(* IEC 61131-3 sources: Industry-PLC-LLM/data/PLCBEAD_repo/PLCBEAD_PLCEmbed-main/PLC-BEAD/Source/PLC_Programs (part 7) *)

(* ---- GEN_RDT.ST ---- *)
FUNCTION _REAL_TO_UDINT:UDINT
  VAR_INPUT
    X :	REAL;
  END_VAR

  IF REAL_TO_UDINT(0.5) = UDINT#1 THEN
    _REAL_TO_UDINT := REAL_TO_UDINT(x);
  ELSIF X > 0.0 THEN
    _REAL_TO_UDINT := REAL_TO_UDINT(x+0.5);
  ELSIF X < 0.0 THEN
    _REAL_TO_UDINT := REAL_TO_UDINT(x-0.5);
  ELSE
    _REAL_TO_UDINT := UDINT#0;
  END_IF;
END_FUNCTION

FUNCTION REAL_TO_TIME2:TIME
	VAR_INPUT
		IN :	REAL;
	END_VAR

	REAL_TO_TIME2 := DINT_TO_TIME(UDINT_TO_DINT(_REAL_TO_UDINT(IN)));
END_FUNCTION

FUNCTION TIME_TO_REAL1:REAL

VAR_INPUT
	X :	TIME;
END_VAR

TIME_TO_REAL1 := UDINT_TO_REAL(DINT_TO_UDINT(TIME_TO_DINT(X)));
END_FUNCTION

FUNCTION D_TRUNC : DINT
  VAR_INPUT
    x : REAL;
  END_VAR

  D_TRUNC := REAL_TO_DINT(X);
  IF X > 0.0 THEN
  	IF DINT_TO_REAL(D_TRUNC) > X THEN D_TRUNC := D_TRUNC - DINT#1; END_IF;
  ELSE
  	IF DINT_TO_REAL(D_TRUNC) < X THEN D_TRUNC := D_TRUNC + DINT#1; END_IF;
  END_IF;
END_FUNCTION

FUNCTION BIT_COUNT:INT

	VAR_INPUT
		IN :	DWORD;
	END_VAR

	VAR
		in_temp :	DWORD;
	END_VAR

	in_temp := IN;
	WHILE in_temp > DWORD#0 DO
		IF (in_temp AND DWORD#16#00000001) > DWORD#0 THEN Bit_Count := Bit_Count +1; END_IF;
		in_temp := SHR(in_temp,1);
	END_WHILE;

END_FUNCTION

FUNCTION FRACT:REAL
	VAR_INPUT
		X :	REAL;
	END_VAR

	IF ABS(x) < 2.0E9 THEN
		FRACT := x - DINT_TO_REAL(D_TRUNC(x));
	ELSE
		FRACT := 0.0;
	END_IF;

END_FUNCTION

FUNCTION_BLOCK T_PLC_MS_block
	VAR_OUTPUT
		T_PLC_MS :	UDINT;
	END_VAR

	VAR_EXTERNAL
		PLC_TICKS_PER_SEC :	INT;
		PLC_SYS_TICK_CNT :	DINT;
	END_VAR

	VAR
		debug :	BOOL;(*Debug-Mode ON / OFF*)
		N :	INT;(*Debug-Faktor*)
		Offset :	UDINT;(*Debug-Offset*)
		temp :	DWORD := DWORD#1;(*Debug-Offset*)
		mode :	BOOL;(*modus*)
		faktor :	UDINT;(*Systemtakt-Faktor*)
		init :	BOOL;
		v_plc_ticks_per_sec :	UDINT;
		base :	UDINT := UDINT#1000;
	END_VAR

	IF init = FALSE THEN
		v_plc_ticks_per_sec := INT_TO_UDINT(PLC_TICKS_PER_SEC);
		IF v_plc_ticks_per_sec = UDINT#1024 THEN
			faktor := UDINT#1;
			mode := FALSE;
		ELSIF v_plc_ticks_per_sec > UDINT#0 THEN
			IF v_plc_ticks_per_sec <= base THEN
				faktor := base / v_plc_ticks_per_sec;
				mode := FALSE;
			ELSE
				faktor := v_plc_ticks_per_sec / base;
				mode := TRUE;
			END_IF;
		ELSE
			faktor := UDINT#1;
		END_IF;
		init := TRUE;
	END_IF;

	IF mode THEN
		T_PLC_MS := DINT_TO_UDINT(PLC_SYS_TICK_CNT) / faktor;
	ELSE
		T_PLC_MS := DINT_TO_UDINT(PLC_SYS_TICK_CNT) * faktor;
	END_IF;

	IF debug THEN
		T_PLC_MS := (DWORD_TO_UDINT(SHL(UDINT_TO_DWORD(T_PLC_MS),N) OR SHL(temp,N)) - UDINT#1) + Offset;
	END_IF;

END_FUNCTION_BLOCK

FUNCTION BIT_LOAD_DW:DWORD

	VAR_INPUT
		IN :	DWORD;
		VAL :	BOOL;
		POS :	INT;
	END_VAR

	IF val THEN
		BIT_LOAD_DW := in OR SHL(DWORD#1,pos);
	ELSE
		BIT_LOAD_DW := in AND (NOT SHL(DWORD#1,pos));
	END_IF;

END_FUNCTION

FUNCTION BIT_OF_DWORD : BOOL
  VAR_INPUT
    IN : DWORD;
    N : INT;
  END_VAR

  BIT_OF_DWORD := (SHR(in,N) AND 16#00000001) > 0;
  (* from OSCAT library; www.oscat.de  *)
END_FUNCTION

FUNCTION _INT_TO_UDINT:UDINT
	VAR_INPUT
		IN :	INT;
	END_VAR

	_INT_TO_UDINT := DINT_TO_UDINT(INT_TO_DINT(IN));
END_FUNCTION

FUNCTION _DWORD_TO_REAL:REAL
	VAR_INPUT
		IN :	DWORD;
	END_VAR

	_DWORD_TO_REAL := UDINT_TO_REAL(DWORD_TO_UDINT(IN));

END_FUNCTION

FUNCTION_BLOCK RDM_block
	VAR_INPUT
		LAST :	REAL;
	END_VAR
	VAR_OUTPUT
		RDM :	REAL;
	END_VAR
	VAR
		T_PLC_MS :	T_PLC_MS_block;
		tn :	DWORD;
		tc :	INT;
	END_VAR
	T_PLC_MS();
	tn := UDINT_TO_DWORD(T_PLC_MS.T_PLC_MS);
	tc := Bit_Count(tn);

	tn:=BIT_LOAD_DW(tn,BIT_OF_DWORD(tn,2),31); (* tn.31 := tn.2; *)
	tn:=BIT_LOAD_DW(tn,BIT_OF_DWORD(tn,5),30); (* tn.30 := tn.5; *)
	tn:=BIT_LOAD_DW(tn,BIT_OF_DWORD(tn,4),29); (* tn.29 := tn.4; *)
	tn:=BIT_LOAD_DW(tn,BIT_OF_DWORD(tn,1),28); (* tn.28 := tn.1; *)
	tn:=BIT_LOAD_DW(tn,BIT_OF_DWORD(tn,0),27); (* tn.27 := tn.0; *)
	tn:=BIT_LOAD_DW(tn,BIT_OF_DWORD(tn,7),26); (* tn.26 := tn.7; *)
	tn:=BIT_LOAD_DW(tn,BIT_OF_DWORD(tn,6),25); (* tn.25 := tn.6; *)
	tn:=BIT_LOAD_DW(tn,BIT_OF_DWORD(tn,3),24); (* tn.24 := tn.3; *)

	tn := ROL(tn,Bit_Count(tn)) OR DWORD#16#80000001;
	tn := UDINT_TO_DWORD(DWORD_TO_UDINT(tn) MOD UDINT#71474513 + _INT_TO_UDINT(tc) + UDINT#77);
	RDM := fract(_DWORD_TO_REAL(tn) / 10000000.0 * (2.71828182845904523536028747135266249 - LIMIT_REAL(0.0,last,1.0)));
END_FUNCTION_BLOCK

FUNCTION_BLOCK GEN_RDT_Block

	VAR_INPUT
		ENABLE :	BOOL := TRUE;
		MIN_TIME_MS :	TIME := t#1s;
		MAX_TIME_MS :	TIME := t#1.2s;
		TP_Q :	TIME := t#100ms;
	END_VAR

	VAR_OUTPUT
		XQ :	BOOL;
	END_VAR

	VAR
		tonRDMTimer :	TON;
		tof_xQ :	TOF;
		tRDMTime :	TIME;
		rRDMTime :	REAL;
		rdm_1 :	RDM_Block;
	END_VAR

	tonRDMTimer(IN:=Enable,PT:=tRDMTime);
	tof_xQ(IN := tonRDMTimer.Q,PT:=TP_Q);
	XQ := tof_xq.Q;
	IF tonRDMTimer.Q THEN
		xQ := TRUE ;
		rdm_1(last:=rRDMTime);
		rRDMTime:= rdm_1.RDM;

		tRDMTime := REAL_TO_TIME2(rRDMTime * TIME_TO_REAL1(Max_Time_ms - Min_Time_ms) + TIME_TO_REAL1(Min_Time_ms));
		tonRDMTimer (IN:=FALSE);
	END_IF;

END_FUNCTION_BLOCK

PROGRAM program0
  VAR
	ENABLE :	BOOL := TRUE;
	MIN_TIME_MS :	TIME := t#1s;
	MAX_TIME_MS :	TIME := t#1.2s;
	TP_Q :	TIME := t#100ms;
	XQ :	BOOL;
	func_block : GEN_RDT_Block;
  END_VAR
	func_block.ENABLE  :=ENABLE;
	func_block.MIN_TIME_MS  :=MIN_TIME_MS;
	func_block.MAX_TIME_MS  :=MAX_TIME_MS;
	func_block.TP_Q  :=TP_Q;
	func_block();
	XQ := func_block.XQ;
END_PROGRAM

CONFIGURATION Config0
	VAR_GLOBAL
		PLC_TICKS_PER_SEC :	INT;
		PLC_SYS_TICK_CNT :	DINT;
	END_VAR
	RESOURCE Res0 ON PLC
		TASK task0(INTERVAL := T#20ms,PRIORITY := 0);
		PROGRAM instance0 WITH task0 : program0;
	END_RESOURCE
END_CONFIGURATION

(* ---- GEN_RMP.ST ---- *)
FUNCTION D_TRUNC : DINT
  VAR_INPUT
    x : REAL;
  END_VAR

  D_TRUNC := REAL_TO_DINT(X);
  IF X > 0.0 THEN
  	IF DINT_TO_REAL(D_TRUNC) > X THEN D_TRUNC := D_TRUNC - DINT#1; END_IF;
  ELSE
  	IF DINT_TO_REAL(D_TRUNC) < X THEN D_TRUNC := D_TRUNC + DINT#1; END_IF;
  END_IF;
END_FUNCTION

FUNCTION FRACT:REAL
	VAR_INPUT
		X :	REAL;
	END_VAR

	IF ABS(x) < 2.0E9 THEN
		FRACT := x - DINT_TO_REAL(D_TRUNC(x));
	ELSE
		FRACT := 0.0;
	END_IF;
END_FUNCTION

FUNCTION _REAL_TO_DWORD: DWORD

  VAR_INPUT
    X :	REAL;
  END_VAR

  IF REAL_TO_DWORD(0.5) = DWORD#1 THEN
    _REAL_TO_DWORD := REAL_TO_DWORD(x);
  ELSIF X > 0.0 THEN
    _REAL_TO_DWORD := REAL_TO_DWORD(x+0.5);
  ELSIF X < 0.0 THEN
    _REAL_TO_DWORD := REAL_TO_DWORD(x-0.5);
  ELSE
    _REAL_TO_DWORD := DWORD#0;
  END_IF;
END_FUNCTION

FUNCTION _DWORD_TO_REAL:REAL
	VAR_INPUT
		IN :	DWORD;
	END_VAR

	_DWORD_TO_REAL := UDINT_TO_REAL(DWORD_TO_UDINT(IN));

END_FUNCTION

FUNCTION MULTIME:TIME
	VAR_INPUT
		T :	TIME;
		M :	REAL;
	END_VAR

	multime := DWORD_TO_TIME(_REAL_TO_DWORD(_DWORD_TO_REAL(TIME_TO_DWORD(t))*M));
END_FUNCTION

FUNCTION TIME_TO_REAL1:REAL

VAR_INPUT
	X :	TIME;
END_VAR

TIME_TO_REAL1 := UDINT_TO_REAL(DINT_TO_UDINT(TIME_TO_DINT(X)));
END_FUNCTION

FUNCTION MODR : REAL
  VAR_INPUT
    IN : REAL;
    DIVI : REAL;
  END_VAR

  IF divi = 0.0 THEN
  	MODR := 0.0;
  ELSE
  	MODR := in - DINT_TO_REAL(FLOOR2(in / divi)) * divi;
  END_IF;
END_FUNCTION

FUNCTION FLOOR2 : DINT
  VAR_INPUT
    x : REAL;
  END_VAR

  FLOOR2 := REAL_TO_DINT(X);
  IF DINT_TO_REAL(FLOOR2) > X THEN
  	FLOOR2 := FLOOR2 - DINT#1;
  END_IF;
END_FUNCTION

FUNCTION UDINT_TO_TIME2:TIME

	VAR_INPUT
		IN :	UDINT;
	END_VAR

	UDINT_TO_TIME2 := DINT_TO_TIME(UDINT_TO_DINT(IN));

END_FUNCTION

FUNCTION_BLOCK T_PLC_MS_block
	VAR_OUTPUT
		T_PLC_MS :	UDINT;
	END_VAR

	VAR_EXTERNAL
		PLC_TICKS_PER_SEC :	INT;
		PLC_SYS_TICK_CNT :	DINT;
	END_VAR

	VAR
		debug :	BOOL;(*Debug-Mode ON / OFF*)
		N :	INT;(*Debug-Faktor*)
		Offset :	UDINT;(*Debug-Offset*)
		temp :	DWORD := DWORD#1;(*Debug-Offset*)
		mode :	BOOL;(*modus*)
		faktor :	UDINT;(*Systemtakt-Faktor*)
		init :	BOOL;
		v_plc_ticks_per_sec :	UDINT;
		base :	UDINT := UDINT#1000;
	END_VAR

	IF init = FALSE THEN
		v_plc_ticks_per_sec := INT_TO_UDINT(PLC_TICKS_PER_SEC);
		IF v_plc_ticks_per_sec = UDINT#1024 THEN
			faktor := UDINT#1;
			mode := FALSE;
		ELSIF v_plc_ticks_per_sec > UDINT#0 THEN
			IF v_plc_ticks_per_sec <= base THEN
				faktor := base / v_plc_ticks_per_sec;
				mode := FALSE;
			ELSE
				faktor := v_plc_ticks_per_sec / base;
				mode := TRUE;
			END_IF;
		ELSE
			faktor := UDINT#1;
		END_IF;
		init := TRUE;
	END_IF;

	IF mode THEN
		T_PLC_MS := DINT_TO_UDINT(PLC_SYS_TICK_CNT) / faktor;
	ELSE
		T_PLC_MS := DINT_TO_UDINT(PLC_SYS_TICK_CNT) * faktor;
	END_IF;

	IF debug THEN
		T_PLC_MS := (DWORD_TO_UDINT(SHL(UDINT_TO_DWORD(T_PLC_MS),N) OR SHL(temp,N)) - UDINT#1) + Offset;
	END_IF;

END_FUNCTION_BLOCK

FUNCTION_BLOCK GEN_RMP_Block

	VAR_INPUT
		PT :	TIME := T#1s;
		AM :	REAL := REAL#1.0;
		OS :	REAL;
		DL :	REAL;
	END_VAR

	VAR_OUTPUT
		Q :	BOOL;
		OUT :	REAL;
	END_VAR

	VAR
		tx :	TIME;
		last :	TIME;
		init :	BOOL;
		temp :	REAL;
		ltemp :	REAL;
		T_PLC_MS :	T_PLC_MS_Block;
	END_VAR

	T_PLC_MS();
	tx:= UDINT_TO_TIME(T_PLC_MS.T_PLC_MS) - last;
	DL := modR(dl,1.0);
	IF dl < 0.0 THEN dl := 1.0 - dl; END_IF;

	IF NOT init THEN
		init := TRUE;
		last := tx;
		tx := t#0s;
	END_IF;

	IF tx >= pt THEN
		last := last + pt;
		tx := tx - pt;
	END_IF;

	ltemp := temp;
	IF pt > t#0s THEN temp := fract(TIME_TO_REAL1(tx + multime(pt, dl)) / TIME_TO_REAL1(pt)); END_IF;
	out := am * temp + os;

	Q := temp < ltemp;

END_FUNCTION_BLOCK

PROGRAM program0
  VAR
	PT :	TIME := T#1s;
	AM :	REAL := REAL#1.0;
	OS :	REAL;
	DL :	REAL;
	Q :	BOOL;
	OUT :	REAL;
	func_block : GEN_RMP_Block;
  END_VAR
	func_block.PT  :=PT;
	func_block.AM  :=AM;
	func_block.OS  :=OS;
	func_block.DL  :=DL;
	func_block();
	Q := func_block.Q;
	OUT := func_block.OUT;
END_PROGRAM

CONFIGURATION Config0
	VAR_GLOBAL
		PLC_TICKS_PER_SEC :	INT;
		PLC_SYS_TICK_CNT :	DINT;
	END_VAR
	RESOURCE Res0 ON PLC
		TASK task0(INTERVAL := T#20ms,PRIORITY := 0);
		PROGRAM instance0 WITH task0 : program0;
	END_RESOURCE
END_CONFIGURATION

(* ---- GEN_SIN.ST ---- *)
FUNCTION _REAL_TO_DWORD: DWORD

  VAR_INPUT
    X :	REAL;
  END_VAR

  IF REAL_TO_DWORD(0.5) = DWORD#1 THEN
    _REAL_TO_DWORD := REAL_TO_DWORD(x);
  ELSIF X > 0.0 THEN
    _REAL_TO_DWORD := REAL_TO_DWORD(x+0.5);
  ELSIF X < 0.0 THEN
    _REAL_TO_DWORD := REAL_TO_DWORD(x-0.5);
  ELSE
    _REAL_TO_DWORD := DWORD#0;
  END_IF;
END_FUNCTION

FUNCTION _DWORD_TO_REAL:REAL
	VAR_INPUT
		IN :	DWORD;
	END_VAR

	_DWORD_TO_REAL := UDINT_TO_REAL(DWORD_TO_UDINT(IN));

END_FUNCTION

FUNCTION MULTIME:TIME
	VAR_INPUT
		T :	TIME;
		M :	REAL;
	END_VAR

	multime := DWORD_TO_TIME(_REAL_TO_DWORD(_DWORD_TO_REAL(TIME_TO_DWORD(t))*M));
END_FUNCTION

FUNCTION UDINT_TO_TIME2:TIME

	VAR_INPUT
		IN :	UDINT;
	END_VAR

	UDINT_TO_TIME2 := DINT_TO_TIME(UDINT_TO_DINT(IN));

END_FUNCTION

FUNCTION_BLOCK T_PLC_MS_block
	VAR_OUTPUT
		T_PLC_MS :	UDINT;
	END_VAR

	VAR_EXTERNAL
		PLC_TICKS_PER_SEC :	INT;
		PLC_SYS_TICK_CNT :	DINT;
	END_VAR

	VAR
		debug :	BOOL;(*Debug-Mode ON / OFF*)
		N :	INT;(*Debug-Faktor*)
		Offset :	UDINT;(*Debug-Offset*)
		temp :	DWORD := DWORD#1;(*Debug-Offset*)
		mode :	BOOL;(*modus*)
		faktor :	UDINT;(*Systemtakt-Faktor*)
		init :	BOOL;
		v_plc_ticks_per_sec :	UDINT;
		base :	UDINT := UDINT#1000;
	END_VAR

	IF init = FALSE THEN
		v_plc_ticks_per_sec := INT_TO_UDINT(PLC_TICKS_PER_SEC);
		IF v_plc_ticks_per_sec = UDINT#1024 THEN
			faktor := UDINT#1;
			mode := FALSE;
		ELSIF v_plc_ticks_per_sec > UDINT#0 THEN
			IF v_plc_ticks_per_sec <= base THEN
				faktor := base / v_plc_ticks_per_sec;
				mode := FALSE;
			ELSE
				faktor := v_plc_ticks_per_sec / base;
				mode := TRUE;
			END_IF;
		ELSE
			faktor := UDINT#1;
		END_IF;
		init := TRUE;
	END_IF;

	IF mode THEN
		T_PLC_MS := DINT_TO_UDINT(PLC_SYS_TICK_CNT) / faktor;
	ELSE
		T_PLC_MS := DINT_TO_UDINT(PLC_SYS_TICK_CNT) * faktor;
	END_IF;

	IF debug THEN
		T_PLC_MS := (DWORD_TO_UDINT(SHL(UDINT_TO_DWORD(T_PLC_MS),N) OR SHL(temp,N)) - UDINT#1) + Offset;
	END_IF;

END_FUNCTION_BLOCK

FUNCTION TIME_TO_REAL1:REAL

	VAR_INPUT
		X :	TIME;
	END_VAR

	TIME_TO_REAL1 := UDINT_TO_REAL(DINT_TO_UDINT(TIME_TO_DINT(X)));
END_FUNCTION

FUNCTION MODR : REAL
  VAR_INPUT
    IN : REAL;
    DIVI : REAL;
  END_VAR

  IF divi = 0.0 THEN
  	MODR := 0.0;
  ELSE
  	MODR := in - DINT_TO_REAL(FLOOR2(in / divi)) * divi;
  END_IF;
END_FUNCTION

FUNCTION FLOOR2 : DINT
  VAR_INPUT
    x : REAL;
  END_VAR

  FLOOR2 := REAL_TO_DINT(X);
  IF DINT_TO_REAL(FLOOR2) > X THEN
  	FLOOR2 := FLOOR2 - DINT#1;
  END_IF;
END_FUNCTION

FUNCTION SIGN_R : BOOL
  VAR_INPUT
    IN : REAL;
  END_VAR

  SIGN_R := in < 0.0;
END_FUNCTION

FUNCTION_BLOCK GEN_SIN_Block

	VAR_INPUT
		PT :	TIME;
		AM :	REAL := REAL#1.0;
		OS :	REAL;
		DL :	REAL;
	END_VAR

	VAR_OUTPUT
		Q :	BOOL;
		Out :	REAL;
	END_VAR

	VAR
		tx :	TIME;
		last :	TIME;
		init :	BOOL;
		temp :	REAL;
		T_PLC_MS :	T_PLC_MS_Block;
	END_VAR

	T_PLC_MS();
	tx:= UDINT_TO_TIME(T_PLC_MS.T_PLC_MS) - last;

	DL := modR(dl,1.0);
	IF dl < 0.0 THEN dl := 1.0 - dl; END_IF;

	IF NOT init THEN
		init := TRUE;
		last := tx;
		tx := t#0s;
	END_IF;

	IF tx >= pt THEN
		last := last + pt;
		tx := tx - pt;
	END_IF;

	IF pt > t#0s THEN temp := SIN(6.283185307179586476 * TIME_TO_REAL1(tx + multime(pt, dl)) / TIME_TO_REAL(pt)); END_IF;
	out := am * 0.5 *  temp + os;

	q := NOT sign_R(temp);

END_FUNCTION_BLOCK

PROGRAM program0
  VAR
	PT :	TIME := T#1s;
	AM :	REAL := REAL#1.0;
	OS :	REAL;
	DL :	REAL;
	Q :	BOOL;
	OUT :	REAL;
	func_block : GEN_SIN_Block;
  END_VAR
	func_block.PT  :=PT;
	func_block.AM  :=AM;
	func_block.OS  :=OS;
	func_block.DL  :=DL;
	func_block();
	Q := func_block.Q;
	OUT := func_block.OUT;
END_PROGRAM

CONFIGURATION Config0
	VAR_GLOBAL
		PLC_TICKS_PER_SEC :	INT;
		PLC_SYS_TICK_CNT :	DINT;
	END_VAR
	RESOURCE Res0 ON PLC
		TASK task0(INTERVAL := T#20ms,PRIORITY := 0);
		PROGRAM instance0 WITH task0 : program0;
	END_RESOURCE
END_CONFIGURATION

(* ---- GEN_SQ.ST ---- *)
FUNCTION UDINT_TO_TIME2:TIME

	VAR_INPUT
		IN :	UDINT;
	END_VAR

	UDINT_TO_TIME2 := DINT_TO_TIME(UDINT_TO_DINT(IN));

END_FUNCTION

FUNCTION_BLOCK T_PLC_MS_block
	VAR_OUTPUT
		T_PLC_MS :	UDINT;
	END_VAR

	VAR_EXTERNAL
		PLC_TICKS_PER_SEC :	INT;
		PLC_SYS_TICK_CNT :	DINT;
	END_VAR

	VAR
		debug :	BOOL;(*Debug-Mode ON / OFF*)
		N :	INT;(*Debug-Faktor*)
		Offset :	UDINT;(*Debug-Offset*)
		temp :	DWORD := DWORD#1;(*Debug-Offset*)
		mode :	BOOL;(*modus*)
		faktor :	UDINT;(*Systemtakt-Faktor*)
		init :	BOOL;
		v_plc_ticks_per_sec :	UDINT;
		base :	UDINT := UDINT#1000;
	END_VAR

	IF init = FALSE THEN
		v_plc_ticks_per_sec := INT_TO_UDINT(PLC_TICKS_PER_SEC);
		IF v_plc_ticks_per_sec = UDINT#1024 THEN
			faktor := UDINT#1;
			mode := FALSE;
		ELSIF v_plc_ticks_per_sec > UDINT#0 THEN
			IF v_plc_ticks_per_sec <= base THEN
				faktor := base / v_plc_ticks_per_sec;
				mode := FALSE;
			ELSE
				faktor := v_plc_ticks_per_sec / base;
				mode := TRUE;
			END_IF;
		ELSE
			faktor := UDINT#1;
		END_IF;
		init := TRUE;
	END_IF;

	IF mode THEN
		T_PLC_MS := DINT_TO_UDINT(PLC_SYS_TICK_CNT) / faktor;
	ELSE
		T_PLC_MS := DINT_TO_UDINT(PLC_SYS_TICK_CNT) * faktor;
	END_IF;

	IF debug THEN
		T_PLC_MS := (DWORD_TO_UDINT(SHL(UDINT_TO_DWORD(T_PLC_MS),N) OR SHL(temp,N)) - UDINT#1) + Offset;
	END_IF;

END_FUNCTION_BLOCK

FUNCTION_BLOCK GEN_SQ_Block

	VAR_INPUT
		PT :	TIME;
	END_VAR

	VAR_OUTPUT
		Q :	BOOL;
	END_VAR

	VAR
		init :	BOOL;
		tn :	TIME;
		tx :	TIME;
		T_PLC_MS :	T_PLC_MS_Block;
	END_VAR

	T_PLC_MS();
	tx := UDINT_TO_TIME(T_PLC_MS.T_PLC_MS);

	IF NOT init THEN
		init := TRUE;
		tn := tx;
		Q := TRUE;
	ELSIF tx - tn >= DWORD_TO_TIME(SHR(TIME_TO_DWORD(PT),1)) THEN
		Q := NOT Q;
		tn := tn + DWORD_TO_TIME(SHR(TIME_TO_DWORD(pt),1));
	END_IF;

END_FUNCTION_BLOCK

PROGRAM program0
  VAR
	PT :	TIME;
	Q :	BOOL;
	OUT :	REAL;
	func_block : GEN_SQ_Block;
  END_VAR
	func_block.PT  :=PT;
	func_block();
	Q := func_block.Q;
END_PROGRAM

CONFIGURATION Config0
	VAR_GLOBAL
		PLC_TICKS_PER_SEC :	INT;
		PLC_SYS_TICK_CNT :	DINT;
	END_VAR
	RESOURCE Res0 ON PLC
		TASK task0(INTERVAL := T#20ms,PRIORITY := 0);
		PROGRAM instance0 WITH task0 : program0;
	END_RESOURCE
END_CONFIGURATION

(* ---- GEN_SQR.ST ---- *)
FUNCTION UDINT_TO_TIME2:TIME

	VAR_INPUT
		IN :	UDINT;
	END_VAR

	UDINT_TO_TIME2 := DINT_TO_TIME(UDINT_TO_DINT(IN));

END_FUNCTION

FUNCTION_BLOCK T_PLC_MS_block
	VAR_OUTPUT
		T_PLC_MS :	UDINT;
	END_VAR

	VAR_EXTERNAL
		PLC_TICKS_PER_SEC :	INT;
		PLC_SYS_TICK_CNT :	DINT;
	END_VAR

	VAR
		debug :	BOOL;(*Debug-Mode ON / OFF*)
		N :	INT;(*Debug-Faktor*)
		Offset :	UDINT;(*Debug-Offset*)
		temp :	DWORD := DWORD#1;(*Debug-Offset*)
		mode :	BOOL;(*modus*)
		faktor :	UDINT;(*Systemtakt-Faktor*)
		init :	BOOL;
		v_plc_ticks_per_sec :	UDINT;
		base :	UDINT := UDINT#1000;
	END_VAR

	IF init = FALSE THEN
		v_plc_ticks_per_sec := INT_TO_UDINT(PLC_TICKS_PER_SEC);
		IF v_plc_ticks_per_sec = UDINT#1024 THEN
			faktor := UDINT#1;
			mode := FALSE;
		ELSIF v_plc_ticks_per_sec > UDINT#0 THEN
			IF v_plc_ticks_per_sec <= base THEN
				faktor := base / v_plc_ticks_per_sec;
				mode := FALSE;
			ELSE
				faktor := v_plc_ticks_per_sec / base;
				mode := TRUE;
			END_IF;
		ELSE
			faktor := UDINT#1;
		END_IF;
		init := TRUE;
	END_IF;

	IF mode THEN
		T_PLC_MS := DINT_TO_UDINT(PLC_SYS_TICK_CNT) / faktor;
	ELSE
		T_PLC_MS := DINT_TO_UDINT(PLC_SYS_TICK_CNT) * faktor;
	END_IF;

	IF debug THEN
		T_PLC_MS := (DWORD_TO_UDINT(SHL(UDINT_TO_DWORD(T_PLC_MS),N) OR SHL(temp,N)) - UDINT#1) + Offset;
	END_IF;

END_FUNCTION_BLOCK

FUNCTION MODR : REAL
  VAR_INPUT
    IN : REAL;
    DIVI : REAL;
  END_VAR

  IF divi = 0.0 THEN
  	MODR := 0.0;
  ELSE
  	MODR := in - DINT_TO_REAL(FLOOR2(in / divi)) * divi;
  END_IF;
END_FUNCTION

FUNCTION FLOOR2 : DINT
  VAR_INPUT
    x : REAL;
  END_VAR

  FLOOR2 := REAL_TO_DINT(X);
  IF DINT_TO_REAL(FLOOR2) > X THEN
  	FLOOR2 := FLOOR2 - DINT#1;
  END_IF;
END_FUNCTION

FUNCTION _REAL_TO_DWORD: DWORD

  VAR_INPUT
    X :	REAL;
  END_VAR

  IF REAL_TO_DWORD(0.5) = DWORD#1 THEN
    _REAL_TO_DWORD := REAL_TO_DWORD(x);
  ELSIF X > 0.0 THEN
    _REAL_TO_DWORD := REAL_TO_DWORD(x+0.5);
  ELSIF X < 0.0 THEN
    _REAL_TO_DWORD := REAL_TO_DWORD(x-0.5);
  ELSE
    _REAL_TO_DWORD := DWORD#0;
  END_IF;
END_FUNCTION

FUNCTION _DWORD_TO_REAL:REAL
	VAR_INPUT
		IN :	DWORD;
	END_VAR

	_DWORD_TO_REAL := UDINT_TO_REAL(DWORD_TO_UDINT(IN));

END_FUNCTION

FUNCTION MULTIME:TIME
	VAR_INPUT
		T :	TIME;
		M :	REAL;
	END_VAR

	multime := DWORD_TO_TIME(_REAL_TO_DWORD(_DWORD_TO_REAL(TIME_TO_DWORD(t))*M));
END_FUNCTION

FUNCTION_BLOCK GEN_SQR_Block

	VAR_INPUT
		PT :	TIME;
		AM :	REAL := REAL#1.0;
		OS :	REAL;
		DC :	REAL := REAL#0.5;
		DL :	REAL;
	END_VAR

	VAR_OUTPUT
		Q :	BOOL;
		Out :	REAL;
	END_VAR

	VAR
		tx :	TIME;
		last :	TIME;
		init :	BOOL;
		T_PLC_MS :	T_PLC_MS_Block;
	END_VAR

	IF dc = 0.0 THEN
		out := -am * 0.5 + os;
		Q := FALSE;
		RETURN;
	ELSIF dc = 1.0 THEN
		out := am * 0.5 + os;
		Q := TRUE;
		RETURN;
	END_IF;

	T_PLC_MS();
	tx:= UDINT_TO_TIME(T_PLC_MS.T_PLC_MS) - last;
	DL := modR(dl,1.0);
	IF dl < 0.0 THEN dl := 1.0 - dl; END_IF;
	dc := modR(dc,1.0);
	IF dc < 0.0 THEN dc := 1.0 - dc; END_IF;

	IF NOT init THEN
		init := TRUE;
		last := tx;
		tx := t#0s;
	END_IF;

	IF tx >= pt THEN
		last := last + pt;
		tx := tx - pt;
	END_IF;

	IF multime(pt, dl + dc) >= pt THEN
		IF tx >= multime(pt, dl + dc - 1.0) THEN
			out := -am * 0.5 + os;
			Q := FALSE;
		END_IF;
		IF tx >= multime(pt, dl) THEN
			out := am * 0.5 + os;
			Q := TRUE;
		END_IF;
	ELSE
		IF tx >= multime(pt, dl) THEN
			out := am * 0.5 + os;
			Q := TRUE;
		END_IF;
		IF tx >= multime(pt, dl + dc) THEN
			out := -am * 0.5 +os;
			Q := FALSE;
		END_IF;
	END_IF;

END_FUNCTION_BLOCK

PROGRAM program0
  VAR
	PT :	TIME;
	AM :	REAL := REAL#1.0;
	OS :	REAL;
	DC :	REAL := REAL#0.5;
	DL :	REAL;
	Q :	BOOL;
	Out :	REAL;
	func_block : GEN_SQR_Block;
  END_VAR
	func_block.PT  :=PT;
	func_block.AM  :=AM;
	func_block.OS  :=OS;
	func_block.DC  :=DC;
	func_block.DL  :=DL;
	func_block();
	Q := func_block.Q;
	OUT := func_block.OUT;
END_PROGRAM

CONFIGURATION Config0
	VAR_GLOBAL
		PLC_TICKS_PER_SEC :	INT;
		PLC_SYS_TICK_CNT :	DINT;
	END_VAR
	RESOURCE Res0 ON PLC
		TASK task0(INTERVAL := T#20ms,PRIORITY := 0);
		PROGRAM instance0 WITH task0 : program0;
	END_RESOURCE
END_CONFIGURATION

(* ---- HEAT_METER.ST ---- *)
FUNCTION UDINT_TO_TIME2:TIME
	VAR_INPUT
		IN :	UDINT;
	END_VAR
	UDINT_TO_TIME2 := DINT_TO_TIME(UDINT_TO_DINT(IN));
END_FUNCTION

FUNCTION_BLOCK T_PLC_MS_block
	VAR_OUTPUT
		T_PLC_MS :	UDINT;
	END_VAR

	VAR_EXTERNAL
		PLC_TICKS_PER_SEC :	INT;
		PLC_SYS_TICK_CNT :	DINT;
	END_VAR

	VAR
		debug :	BOOL;(*Debug-Mode ON / OFF*)
		N :	INT;(*Debug-Faktor*)
		Offset :	UDINT;(*Debug-Offset*)
		temp :	DWORD := DWORD#1;(*Debug-Offset*)
		mode :	BOOL;(*modus*)
		faktor :	UDINT;(*Systemtakt-Faktor*)
		init :	BOOL;
		v_plc_ticks_per_sec :	UDINT;
		base :	UDINT := UDINT#1000;
	END_VAR

	IF init = FALSE THEN
		v_plc_ticks_per_sec := INT_TO_UDINT(PLC_TICKS_PER_SEC);
		IF v_plc_ticks_per_sec = UDINT#1024 THEN
			faktor := UDINT#1;
			mode := FALSE;
		ELSIF v_plc_ticks_per_sec > UDINT#0 THEN
			IF v_plc_ticks_per_sec <= base THEN
				faktor := base / v_plc_ticks_per_sec;
				mode := FALSE;
			ELSE
				faktor := v_plc_ticks_per_sec / base;
				mode := TRUE;
			END_IF;
		ELSE
			faktor := UDINT#1;
		END_IF;
		init := TRUE;
	END_IF;

	IF mode THEN
		T_PLC_MS := DINT_TO_UDINT(PLC_SYS_TICK_CNT) / faktor;
	ELSE
		T_PLC_MS := DINT_TO_UDINT(PLC_SYS_TICK_CNT) * faktor;
	END_IF;

	IF debug THEN
		T_PLC_MS := (DWORD_TO_UDINT(SHL(UDINT_TO_DWORD(T_PLC_MS),N) OR SHL(temp,N)) - UDINT#1) + Offset;
	END_IF;

END_FUNCTION_BLOCK

TYPE
	oscat_ARRAY_X               : ARRAY [0..1]    OF REAL;
	oscat_XY                    : ARRAY [1..20]   OF oscat_ARRAY_X := [0,0,0,0,0,0,0,0,0,0,0,0,0,0,0,0,0,0,0,0];
END_TYPE

FUNCTION_BLOCK LINEAR_INT_Block

	VAR_INPUT
		X :	REAL;
		XY :	oscat_XY;
		PTS :	INT;
	END_VAR

	VAR_OUTPUT
		LINEAR_INT :	REAL;
	END_VAR

	VAR
		i :	INT;
		i2 :	INT;
	END_VAR

	pts := MIN(pts,20);

	i := 2;

	WHILE (i < pts) AND (XY[i][0] < X) DO
		i := i + 1;
	END_WHILE;

	i2 := i-1;

	LINEAR_INT := ((XY[i][1] - XY[i2][1]) * X - XY[i][1] * XY[i2][0] + XY[i2][1] * XY[i][0]) / (XY[i][0] - XY[i2][0]);

END_FUNCTION_BLOCK

FUNCTION_BLOCK WATER_ENTHALPY_Block

    VAR_INPUT
        T :	REAL;
    END_VAR

    VAR_OUTPUT
        RESULT :	REAL;
    END_VAR

    VAR
        Pts :	INT;
        data :	oscat_XY;
        FB_LINEAR_INT :	LINEAR_INT_Block;
    END_VAR

    IF Pts = 0 THEN
        Pts := 11;
        data[01][0] := REAL#0.0;
        data[01][1] := REAL#0.06;
        data[02][0] := REAL#10.0;
        data[02][1] := REAL#42.1;
        data[03][0] := REAL#20.0;
        data[03][1] := REAL#83.9;
        data[04][0] := REAL#30.0;
        data[04][1] := REAL#125.8;
        data[05][0] := REAL#40.0;
        data[05][1] := REAL#167.58;
        data[06][0] := REAL#50.0;
        data[06][1] := REAL#209.4;
        data[07][0] := REAL#60.0;
        data[07][1] := REAL#251.2;
        data[08][0] := REAL#70.0;
        data[08][1] := REAL#293.1;
        data[09][0] := REAL#80.0;
        data[09][1] := REAL#335.0;
        data[10][0] := REAL#90.0;
        data[10][1] := REAL#377.0;
        data[11][0] := REAL#100.0;
        data[11][1] := REAL#419.1;
    END_IF;

    FB_LINEAR_INT(X:=T,XY:=Data,Pts:=Pts);
    Result :=FB_LINEAR_INT.LINEAR_INT;

END_FUNCTION_BLOCK

FUNCTION_BLOCK R2_SET_Block

	VAR_INPUT
		X :	REAL;
	END_VAR

	VAR_OUTPUT
		R2_SET :	REAL2;
	END_VAR

	R2_SET.RX := X;
	R2_SET.R1 := 0.0;

END_FUNCTION_BLOCK

FUNCTION_BLOCK R2_ADD_Block

	VAR_INPUT
		X :	REAL2;
		Y :	REAL;
	END_VAR

	VAR_OUTPUT
		R2_ADD :	REAL2;
	END_VAR

	VAR
		temp :	REAL;
	END_VAR

	temp := X.RX;
	R2_ADD.RX := Y + X.R1 + X.RX;
	R2_ADD.R1 := temp - R2_ADD.RX + Y + X.R1;

END_FUNCTION_BLOCK

TYPE REAL2:

	STRUCT
		R1 : REAL;
		RX : REAL;
	END_STRUCT;

END_TYPE

FUNCTION_BLOCK INTEGRATE

	VAR_INPUT
		E :	BOOL := TRUE;
		X :	REAL;
		K :	REAL := 1.0;
	END_VAR

	VAR_IN_OUT
		Y :	REAL;
	END_VAR

	VAR
		X_last :	REAL;
		init :	BOOL;
		T_PLC_MS :	T_PLC_MS_block;
		last :	UDINT;
		tx :	UDINT;
	END_VAR

	T_PLC_MS();
	tx:= T_PLC_MS.T_PLC_MS;

	IF NOT init THEN
		init := TRUE;
		X_last := X;
	ELSIF E THEN
		Y := (X + X_LAST) * 0.5E-3 * UDINT_TO_REAL(tx-last) * K + Y;
		X_last := X;
	END_IF;
	last := tx;

END_FUNCTION_BLOCK

FUNCTION_BLOCK FT_INT2_Block

	VAR_INPUT
		IN :	REAL;
		K :	REAL := 1.0;
		RUN :	BOOL := TRUE;
		RST :	BOOL;
		OUT_MIN :	REAL := REAL#-1.0E-37;
		OUT_MAX :	REAL := REAL#1.0E37;
	END_VAR

	VAR_OUTPUT
		OUT :	REAL;
		LIM :	BOOL;
	END_VAR

	VAR
		integ :	INTEGRATE;
		ix :	REAL;
		val :	REAL2;
		R2_ADD :	R2_ADD_Block;
		R2_SET :	R2_SET_Block;
	END_VAR

	IF RST THEN
		R2_SET(X:=0.0);
		val:=R2_SET.R2_SET;
		out := 0.0;
	ELSE
		integ(X := IN, E := RUN, K := K, Y := ix);
		ix := integ.Y;
		R2_ADD(X:=val,Y:=ix);
		val:=R2_ADD.R2_ADD;
		ix := 0.0;
		OUT := val.RX;
	END_IF;

	(* check output for limits *)
	IF out > OUT_MIN AND out < OUT_MAX THEN
		LIM := FALSE;
	ELSE
		OUT := LIMIT(OUT_MIN, OUT, OUT_MAX);
		R2_SET(X:=OUT);
		val:=R2_SET.R2_SET;
		LIM := TRUE;
	END_IF;

END_FUNCTION_BLOCK

FUNCTION WATER_DENSITY:REAL

    VAR_INPUT
        T :	REAL;
        SAT :	BOOL;
    END_VAR

    VAR
        T2 :	REAL;
        T4 :	REAL;
    END_VAR

    T2 := T * T;
    T4 := T2 * T2;
    WATER_DENSITY := (999.83952 + 16.952577*T + -7.9905127E-3*T2 + -4.6241757E-5*T2*T + 1.0584601E-7*T4 + -2.8103006E-10*T4*T) / (1.0 + 0.0168872*T);
    IF sat THEN WATER_DENSITY := WATER_DENSITY - 0.004612 + 0.000106 * T; END_IF;

END_FUNCTION

FUNCTION TIME_TO_UDINT2:UDINT
	VAR_INPUT
		X :	TIME;
	END_VAR

	TIME_TO_UDINT2 := DINT_TO_UDINT(TIME_TO_DINT(X));
END_FUNCTION

FUNCTION_BLOCK HEAT_METER_Block

	VAR_INPUT
		TF :	REAL;
		TR :	REAL;
		LPH :	REAL;
		E :	BOOL;
		RST :	BOOL;
		CP :	REAL;
		DENSITY :	REAL;
		CONTENT :	REAL;
		PULSE_MODE :	BOOL;
		RETURN_METER :	BOOL;
		AVG_TIME :	TIME := T#5s;
	END_VAR

	VAR_OUTPUT
		C :	REAL;
	END_VAR

	VAR_IN_OUT
		Y :	REAL;
	END_VAR

	VAR
		tx :	UDINT;
		last :	UDINT;
		int1 :	FT_INT2_Block;
		edge :	BOOL;
		x :	REAL;
		init :	BOOL;
		Y_last :	REAL;
		T_PLC_MS :	T_PLC_MS_Block;
		WATER_ENTHALPY :	WATER_ENTHALPY_Block;
		wa_TF :	REAL;
		wa_TR :	REAL;
	END_VAR

	IF rst THEN
		int1(rst := TRUE);
		int1.rst := FALSE;
		C := 0.0;
		Y := 0.0;
	ELSIF e THEN
		water_enthalpy(T:=TF);
		wa_TF:=water_enthalpy.Result;

		water_enthalpy(T:=TR);
		wa_TR:=water_enthalpy.Result;

		X := (WATER_DENSITY(SEL(return_meter, TF, TR), FALSE) * (wa_TF - wa_TR) * (1.0 - content) + CP * Density * content * (TF-TR));
	END_IF;

	int1(run := NOT pulse_mode AND e, in := X * LPH * 2.77777777777E-4);
	IF pulse_mode THEN
		IF NOT edge AND E THEN Y := Y + X * LPH; END_IF;
	ELSE
		Y := int1.Out;
	END_IF;

	edge := e;

	T_PLC_MS();
	tx:= T_PLC_MS.T_PLC_MS;

	IF NOT init THEN
		init := TRUE;
		last := tx;
	END_IF;

	IF (tx - last >= TIME_TO_UDINT2(AVG_TIME)) AND (avg_time > T#0s) THEN
		last := tx;
		C := (Y - Y_last) * 3.6E12 / TIME_TO_REAL(AVG_TIME);
		Y_last := Y;
	END_IF;

END_FUNCTION_BLOCK

PROGRAM program0
	VAR
	    TF :	REAL;
		TR :	REAL;
		LPH :	REAL;
		E :	BOOL;
		RST :	BOOL;
		CP :	REAL;
		DENSITY :	REAL;
		CONTENT :	REAL;
		PULSE_MODE :	BOOL;
		RETURN_METER :	BOOL;
		AVG_TIME :	TIME := T#5s;
		Y :	REAL;
		C :	REAL;

		func_block : HEAT_METER_Block;
  	END_VAR
	func_block.TF := TF;
	func_block.TR := TR;
	func_block.LPH := LPH;
	func_block.E := E;
	func_block.RST := RST;
	func_block.CP := CP;
	func_block.DENSITY := DENSITY;
	func_block.CONTENT := CONTENT;
	func_block.PULSE_MODE := PULSE_MODE;
	func_block.RETURN_METER := RETURN_METER;
	func_block.AVG_TIME := AVG_TIME;
	func_block.Y := Y;

	func_block();
	Y := func_block.Y;
	C := func_block.C;
END_PROGRAM

CONFIGURATION Config0
	VAR_GLOBAL
		PLC_TICKS_PER_SEC :	INT;
		PLC_SYS_TICK_CNT :	DINT;
	END_VAR
  	RESOURCE Res0 ON PLC
    	TASK task0(INTERVAL := T#20ms,PRIORITY := 0);
    	PROGRAM instance0 WITH task0 : program0;
  	END_RESOURCE
END_CONFIGURATION

(* ---- HEAT_TEMP.ST ---- *)
FUNCTION_BLOCK HEAT_TEMP_Block

	VAR_INPUT
		T_EXT :	REAL;
		T_INT :	REAL;
		OFFSET :	REAL;
		T_REQ :	REAL;
		TY_MAX :	REAL := REAL#70.0;
		TY_MIN :	REAL := REAL#25.0;
		TY_CONFIG :	REAL := REAL#70.0;
		T_INT_CONFIG :	REAL := REAL#20.0;
		T_EXT_CONFIG :	REAL := REAL#-15.0;
		T_DIFF :	REAL := REAL#10.0;
		C :	REAL := REAL#1.33;
		H :	REAL := REAL#3.0;
	END_VAR

	VAR_OUTPUT
		TY :	REAL;
		HEAT :	BOOL;
	END_VAR

	VAR
		tr :	REAL;
		tx :	REAL;
	END_VAR

	tr := T_INT + OFFSET;
	tx := (tr - T_EXT) / (T_INT_CONFIG - T_EXT_CONFIG);

	IF T_EXT + H > tr THEN
		TY := 0.0;
	ELSE
		TY := LIMIT(TY_MIN, tr + T_DIFF * 0.5 * tx + (TY_CONFIG - T_DIFF * 0.5 - tr) * EXPT(tx, 1.0 / C), TY_MAX);
	END_IF;

	TY := MAX(TY, T_REQ);
	HEAT := TY > 0.0;

END_FUNCTION_BLOCK

PROGRAM program0
	VAR
		T_EXT :	REAL;
		T_INT :	REAL;
		OFFSET :	REAL;
		T_REQ :	REAL;
		TY_MAX :	REAL := REAL#70.0;
		TY_MIN :	REAL := REAL#25.0;
		TY_CONFIG :	REAL := REAL#70.0;
		T_INT_CONFIG :	REAL := REAL#20.0;
		T_EXT_CONFIG :	REAL := REAL#-15.0;
		T_DIFF :	REAL := REAL#10.0;
		C :	REAL := REAL#1.33;
		H :	REAL := REAL#3.0;
		TY :	REAL;
		HEAT :	BOOL;

		func_block : HEAT_TEMP_Block;
	END_VAR
	func_block.T_EXT := T_EXT;
	func_block.T_INT := T_INT;
	func_block.OFFSET := OFFSET ;
	func_block.T_REQ    := T_REQ    ;
	func_block.TY_MAX := TY_MAX;
	func_block.TY_MIN := TY_MIN;
	func_block.TY_CONFIG := TY_CONFIG ;
	func_block.T_INT_CONFIG := T_INT_CONFIG ;
	func_block.T_EXT_CONFIG    := T_EXT_CONFIG    ;
	func_block.T_DIFF    := T_DIFF    ;
	func_block.C := C;
	func_block.H := H;

	func_block();
	TY  := func_block.TY;
	HEAT  := func_block.HEAT;
END_PROGRAM

CONFIGURATION Config0
	RESOURCE Res0 ON PLC
		TASK task0(INTERVAL := T#20ms,PRIORITY := 0);
		PROGRAM instance0 WITH task0 : program0;
	END_RESOURCE
END_CONFIGURATION

(* ---- HEX_TO_BYTE.ST ---- *)
TYPE
	 oscat_STRING5  : STRING;
END_TYPE

FUNCTION_BLOCK HEX_TO_BYTE_Block

	VAR_INPUT
		HEX :	oscat_STRING5;
	END_VAR

	VAR_OUTPUT
		HEX_TO_BYTE :	BYTE;
	END_VAR

	VAR
		i :	INT;
		stop :	INT;
		X :	INT;
	END_VAR

	HEX_TO_BYTE := BYTE#0;
	stop := LEN(HEX);
	FOR I := 1 TO stop DO
		x := GET_CHAR(Hex,I);
		IF X > 47 AND x < 58 THEN
			HEX_TO_BYTE := SHL(HEX_TO_BYTE,4) OR INT_TO_BYTE (X - 48);
		ELSIF X > 64 AND X < 71 THEN
			HEX_TO_BYTE := SHL(HEX_TO_BYTE,4) OR INT_TO_BYTE (X - 55);
		ELSIF X > 96 AND X < 103 THEN
			HEX_TO_BYTE := SHL(HEX_TO_BYTE,4) OR INT_TO_BYTE (X - 87);
		END_IF;
	END_FOR;

END_FUNCTION_BLOCK

PROGRAM program0
  VAR
	HEX :	oscat_STRING5;
	HEX_TO_BYTE :	BYTE;
	func_block : HEX_TO_BYTE_Block;
  END_VAR
	func_block.HEX  :=HEX;
	func_block();
	HEX_TO_BYTE := func_block.HEX_TO_BYTE;
END_PROGRAM

CONFIGURATION Config0
	RESOURCE Res0 ON PLC
		TASK task0(INTERVAL := T#20ms,PRIORITY := 0);
		PROGRAM instance0 WITH task0 : program0;
	END_RESOURCE
END_CONFIGURATION

(* ---- HEX_TO_DWORD.ST ---- *)
FUNCTION_BLOCK HEX_TO_DWORD

	VAR_INPUT
		HEX :	oscat_STRING20;
	END_VAR

	VAR_OUTPUT
		HEX_TO_DWORD :	DWORD;
	END_VAR

	VAR
		i :	INT;
		stop :	INT;
		X :	INT;
	END_VAR

	HEX_TO_DWORD := DWORD#0;
	stop := LEN(Hex);
	FOR I := 1 TO stop DO
		x := GET_CHAR(Hex,I);
		IF X > 47 AND x < 58 THEN
			HEX_TO_DWORD := SHL_DWORD(HEX_TO_DWORD,4) OR INT_TO_DWORD (X - 48);
		ELSIF X > 64 AND X < 71 THEN
			HEX_TO_DWORD := SHL_DWORD(HEX_TO_DWORD,4) OR INT_TO_DWORD (X - 55);
		ELSIF X > 96 AND X < 103 THEN
			HEX_TO_DWORD := SHL_DWORD(HEX_TO_DWORD,4) OR INT_TO_DWORD (X - 87);
		END_IF;
	END_FOR;

END_FUNCTION_BLOCK

(* ---- HOLIDAY.ST ---- *)
TYPE oscat_LANGUAGE:
  STRUCT
    DEFAULT 	: INT;
	LMAX    	: INT;
  END_STRUCT;
END_TYPE

TYPE
	oscat_LOCATION_ELEMENTS	: ARRAY [1..5] OF INT;
END_TYPE

TYPE
  oscat_ELEMENT_WEEKDAYS	: ARRAY [1..7] OF STRING;
  oscat_WEEKDAYS			: ARRAY [1..3]  OF oscat_ELEMENT_WEEKDAYS := [0, 0, 0];
END_TYPE

TYPE oscat_LOCATION:
  STRUCT
    DEFAULT 	: INT;
	LMAX    	: INT;
	LANGUAGE	: oscat_LOCATION_ELEMENTS;
  END_STRUCT;
END_TYPE

TYPE oscat_HOLIDAY_DATA :
  STRUCT
	NAME : STRING;
	DAY : SINT;
	MONTH : SINT;
	USE : SINT;
	PAD_BYTE : BYTE;
  END_STRUCT;
END_TYPE

TYPE
  oscat_HOLIDAY_DATA_0_29 	: ARRAY [0..29] OF oscat_HOLIDAY_DATA;
  oscat_HOLIDAY_DATA_0_49 	: ARRAY [0..49] OF oscat_HOLIDAY_DATA;
END_TYPE

FUNCTION_BLOCK SETUP_LANGUAGE_Block

	VAR_IN_OUT
		LANGUAGE :	oscat_LANGUAGE;
	END_VAR

	VAR
		init :	BOOL;
	END_VAR

	IF init THEN RETURN; END_IF;
	init := TRUE;

	LANGUAGE.DEFAULT  := 1; (* 1=english, 2=german 3=french *)
	LANGUAGE.LMAX := 3;
END_FUNCTION_BLOCK

FUNCTION_BLOCK SETUP_LOCATION
	VAR_IN_OUT
		LOCATION :	oscat_LOCATION;
	END_VAR

	VAR
		init :	BOOL;
	END_VAR

	IF init THEN RETURN; END_IF;
	init := TRUE;

	LOCATION.DEFAULT  := 1;
	LOCATION.LMAX := 5;

	LOCATION.LANGUAGE[1] := 2;
	LOCATION.LANGUAGE[2] := 2;
	LOCATION.LANGUAGE[3] := 3;
	LOCATION.LANGUAGE[4] := 2;
	LOCATION.LANGUAGE[5] := 2;
END_FUNCTION_BLOCK

FUNCTION_BLOCK SETUP_WEEKDAYS

	VAR_IN_OUT
		WEEKDAYS :	oscat_WEEKDAYS;
	END_VAR

	VAR
		init :	BOOL;
	END_VAR

	IF init THEN RETURN; END_IF;
	init := TRUE;

	WEEKDAYS[1][01] := 'Monday';
	WEEKDAYS[1][02] := 'Tuesday';
	WEEKDAYS[1][03] := 'Wednesday';
	WEEKDAYS[1][04] := 'Thursday';
	WEEKDAYS[1][05] := 'Friday';
	WEEKDAYS[1][06] := 'Saturday';
	WEEKDAYS[1][07] := 'Sunday';

	WEEKDAYS[2][01] := 'Montag';
	WEEKDAYS[2][02] := 'Dienstag';
	WEEKDAYS[2][03] := 'Mittwoch';
	WEEKDAYS[2][04] := 'Donnerstag';
	WEEKDAYS[2][05] := 'Freitag';
	WEEKDAYS[2][06] := 'Samstag';
	WEEKDAYS[2][07] := 'Sonntag';

	WEEKDAYS[3][01] := 'Lundi';
	WEEKDAYS[3][02] := 'Mardi';
	WEEKDAYS[3][03] := 'Mercredi';
	WEEKDAYS[3][04] := 'Jeudi';
	WEEKDAYS[3][05] := 'Vendredi';
	WEEKDAYS[3][06] := 'Samedi';
	WEEKDAYS[3][07] := 'Dimanche';
END_FUNCTION_BLOCK

FUNCTION YEAR_OF_DATE:INT
	VAR_INPUT
		IDATE :	UDINT;
	END_VAR

	YEAR_OF_DATE := UDINT_TO_INT((idate+UDINT#43200) / UDINT#31557600 + UDINT#1970);
END_FUNCTION

FUNCTION _INT_TO_UDINT:UDINT
	VAR_INPUT
		IN :	INT;
	END_VAR

	_INT_TO_UDINT := DINT_TO_UDINT(INT_TO_DINT(IN));
END_FUNCTION

FUNCTION SET_DATE:UDINT

	VAR_INPUT
		YEAR :	INT;
		MONTH :	INT;
		DAY :	INT;
	END_VAR

	VAR
		count :	INT;
	END_VAR

	IF month > 2 THEN
		count := (month - 1) * 30;
		IF month > 7 THEN
			count := count + DWORD_TO_INT(SHR(DINT_TO_DWORD(INT_TO_DINT(month) - INT_TO_DINT(3)),1));
		ELSE
			count := count + DWORD_TO_INT(SHR(DINT_TO_DWORD(INT_TO_DINT(month) - INT_TO_DINT(4)),1));
		END_IF;
		IF SHL(INT_TO_WORD(year),14) = WORD#0 THEN
			count := count + 1;
		END_IF;
	ELSE
		count := (month - 1) * 31;
	END_IF;
	SET_DATE := (_INT_TO_UDINT(count + day - 1) + DWORD_TO_UDINT(SHR(UDINT_TO_DWORD(_INT_TO_UDINT(year) * UDINT#1461 - UDINT#2878169), 2))) * UDINT#86400;
END_FUNCTION

FUNCTION DAY_OF_WEEK:INT
	VAR_INPUT
		IDATE :	UDINT;
	END_VAR

	DAY_OF_WEEK := UDINT_TO_INT((idate / UDINT#86400 + UDINT#3) MOD UDINT#7) + INT#01;
END_FUNCTION

FUNCTION EASTER:UDINT
	VAR_INPUT
		YEAR :	INT;
	END_VAR

	VAR
		b :	INT;
		c :	INT;
		oday :	INT;
	END_VAR

	b := (204 - 11 * (year MOD 19)) MOD 30;
	IF b > 27 THEN b := b - 1; END_IF;
	c := (year + WORD_TO_INT(SHR(INT_TO_WORD(year),2)) + b - 13) MOD 7;
	oday := 28 + b - c;
	IF oday > 33 THEN
		easter := set_Date(year, 4, oday - 31);
	ELSE
		easter := set_Date(year, 3, oday);
	END_IF;
END_FUNCTION

FUNCTION LEAP_OF_DATE:BOOL

	VAR_INPUT
		IDATE :	UDINT;
	END_VAR

	LEAP_OF_DATE := SHL(UDINT_TO_DWORD((idate + UDINT#43200) / UDINT#31557600), 30) = DWORD#16#80000000;
END_FUNCTION

FUNCTION DAY_OF_YEAR:INT
	VAR_INPUT
		IDATE :	UDINT;
	END_VAR

	DAY_OF_YEAR := UDINT_TO_INT(((idate) / UDINT#86400) MOD UDINT#1461);
	IF DAY_OF_YEAR > 729 THEN
		IF DAY_OF_YEAR > 1095 THEN DAY_OF_YEAR := DAY_OF_YEAR - 1095; ELSE DAY_OF_YEAR := DAY_OF_YEAR - 729; END_IF;
	ELSIF DAY_OF_YEAR > 364 THEN
		DAY_OF_YEAR := DAY_OF_YEAR - 364;
	ELSE
		DAY_OF_YEAR := DAY_OF_YEAR + 1;
	END_IF;
END_FUNCTION

FUNCTION MONTH_OF_DATE:INT

	VAR_INPUT
		IDATE :	UDINT;
	END_VAR

	MONTH_OF_DATE := DAY_OF_YEAR(idate);
	IF MONTH_OF_DATE < 32 THEN
		MONTH_OF_DATE := 1;
	ELSIF LEAP_OF_DATE((IDATE)) THEN
		MONTH_OF_DATE := (MONTH_OF_DATE * 53 + 1668) / 1623;
	ELSE
		MONTH_OF_DATE := (MONTH_OF_DATE * 53 + 1700) / 1620;
	END_IF;
END_FUNCTION

FUNCTION DAY_OF_MONTH:INT
	VAR_INPUT
		IDATE :	UDINT;
	END_VAR

	day_of_month := day_of_year(idate);

	IF leap_of_Date((idate)) THEN
		CASE day_of_month OF
			32..60	:	day_of_month := day_of_month - 31;
			61..91	:	day_of_month := day_of_month - 60;
			92..121 :	day_of_month := day_of_month - 91;
			122..152:	day_of_month := day_of_month - 121;
			153..182:	day_of_month := day_of_month - 152;
			183..213:	day_of_month := day_of_month - 182;
			214..244:	day_of_month := day_of_month - 213;
			245..274:	day_of_month := day_of_month - 244;
			275..305:	day_of_month := day_of_month - 274;
			306..335:	day_of_month := day_of_month - 305;
			336..366:	day_of_month := day_of_month - 335;
		END_CASE;
	ELSE
		CASE day_of_month OF
			32..59	:	day_of_month := day_of_month - 31;
			60..90	:	day_of_month := day_of_month - 59;
			91..120 :	day_of_month := day_of_month - 90;
			121..151:	day_of_month := day_of_month - 120;
			152..181:	day_of_month := day_of_month - 151;
			182..212:	day_of_month := day_of_month - 181;
			213..243:	day_of_month := day_of_month - 212;
			244..273:	day_of_month := day_of_month - 243;
			274..304:	day_of_month := day_of_month - 273;
			305..334:	day_of_month := day_of_month - 304;
			335..365:	day_of_month := day_of_month - 334;
		END_CASE;
	END_IF;
END_FUNCTION

FUNCTION DATE_ADD:UDINT
	VAR_INPUT
		IDATE :	UDINT;
		D :	INT;
		W :	INT;
		M :	INT;
		Y :	INT;
	END_VAR

	VAR
		mo :	INT;
		yr :	INT;
		dm :	INT;
	END_VAR

	DATE_ADD := IDATE + INT_TO_UDINT(D + W * 7) * UDINT#86400;
	yr := Y + YEAR_OF_DATE(DATE_ADD);
	mo := M + MONTH_OF_DATE(DATE_ADD);
	dm := DAY_OF_MONTH(DATE_ADD);
	WHILE mo > 12 DO
		mo := mo - 12;
		yr := yr + 1;
	END_WHILE;
	WHILE mo < 1 DO
		mo := mo + 12;
		yr := yr - 1;
	END_WHILE;
	DATE_ADD := SET_DATE(yr, mo, dm);
END_FUNCTION

FUNCTION_BLOCK HOLIDAY_Block
	VAR_INPUT
		DATE_IN :	UDINT;
		LANGU :	INT;
		FRIDAY :	BOOL;
		SATURDAY :	BOOL;
		SUNDAY :	BOOL;
	END_VAR

	VAR_IN_OUT
		HOLIDAYS :	oscat_HOLIDAY_DATA_0_29;
	END_VAR

	VAR_OUTPUT
		Y :	BOOL;
		NAME :	STRING;
	END_VAR

	VAR
		size :	INT := INT#29;
		last_active :	UDINT;
		ostern :	UDINT;
		i :	INT;
		jahr :	INT;
		x_date :	UDINT;
		lx :	INT;
		wdx :	INT;
		SETUP_LOCATIONS :	SETUP_LOCATION;
		SETUP_WEEKDAYSS :	SETUP_WEEKDAYS;
		SETUP_LANGUAGES :	SETUP_LANGUAGE_Block;
		LOCATION :	oscat_LOCATION;
		WEEKDAYS :	oscat_WEEKDAYS;
		LANGUAGE :	oscat_LANGUAGE;
		wd :	INT;
	END_VAR

	IF last_active = date_in THEN RETURN; END_IF;
	last_active := DATE_IN;

	SETUP_LOCATIONS(LOCATION:=LOCATION);
	LOCATION:=SETUP_LOCATIONS.LOCATION;

	SETUP_WEEKDAYSS(WEEKDAYS:=WEEKDAYS);
	WEEKDAYS:=SETUP_WEEKDAYSS.WEEKDAYS;

	SETUP_LANGUAGES(LANGUAGE:=LANGUAGE);
	LANGUAGE:=SETUP_LANGUAGES.LANGUAGE;

	IF LANGU = 0 THEN
		lx := language.DEFAULT;
	ELSE
		lx := MIN(language.LMAX, LANGU);
	END_IF;

	jahr := YEAR_OF_DATE(date_in);
	ostern := EASTER(jahr);
	wdx := DAY_OF_WEEK(DATE_IN);
	Y := FALSE;

	FOR i := 0 TO size DO
		x_date := SET_DATE(jahr, SINT_TO_INT(HOLIDAYS[i].MONTH) , SINT_TO_INT(HOLIDAYS[i].DAY));
		IF HOLIDAYS[i].USE = SINT#1 AND HOLIDAYS[i].MONTH > SINT#0 THEN
			(* check for fixed date holiday *)
			IF x_date = date_in THEN
				Y := TRUE;
				NAME := HOLIDAYS[i].NAME;
				RETURN;
			END_IF;
		ELSIF HOLIDAYS[i].USE = SINT#1 AND HOLIDAYS[i].MONTH = SINT#0 THEN
			(* check for holiday in reference to easter *)
			IF DATE_ADD(ostern, SINT_TO_INT(HOLIDAYS[i].DAY),0,0,0) = date_in THEN
				Y := TRUE;
				NAME := HOLIDAYS[i].NAME;
				RETURN;
			END_IF;
		ELSIF HOLIDAYS[i].USE < SINT#0 THEN
			(* check for holiday on a weekday before date *)
			IF DAY_OF_WEEK(date_in) = SINT_TO_INT(ABS(HOLIDAYS[i].USE)) AND date_in < x_date AND date_in >= DATE_ADD(x_date,-7,0,0,0) THEN
				Y := TRUE;
				NAME := HOLIDAYS[i].NAME;
				RETURN;
			END_IF;
		END_IF;
	END_FOR;

	IF NOT Y AND (wdx = 5 AND FRIDAY OR wdx = 6 AND SATURDAY OR wdx = 7 AND SUNDAY) THEN
		Y := TRUE;
		wd := LOCATION.LANGUAGE[lx];
		NAME := WEEKDAYS[wd][wdx];
	ELSE
		NAME := '';
	END_IF;
END_FUNCTION_BLOCK

PROGRAM program0
  VAR
	DATE_IN  :	UDINT;
	LANGU    :	INT;
	FRIDAY   :	BOOL;
	SATURDAY :	BOOL;
	SUNDAY   :	BOOL;

	Y :	BOOL;
	NAME :	STRING;

	HOLIDAYS :	oscat_HOLIDAY_DATA_0_29;

	func_block : HOLIDAY_Block;
  END_VAR
	func_block.DATE_IN :=DATE_IN ;
	func_block.LANGU   :=LANGU   ;
	func_block.FRIDAY  :=FRIDAY  ;
	func_block.SATURDAY:=SATURDAY;
	func_block.SUNDAY  :=SUNDAY  ;
	func_block.HOLIDAYS  :=HOLIDAYS ;

	func_block();
	Y := func_block.Y;
	NAME := func_block.NAME;
	HOLIDAYS := func_block.HOLIDAYS;

END_PROGRAM

CONFIGURATION Config0
  RESOURCE Res0 ON PLC
    TASK task0(INTERVAL := T#20ms,PRIORITY := 0);
    PROGRAM instance0 WITH task0 : program0;
  END_RESOURCE
END_CONFIGURATION

(* ---- HTML_DECODE.ST ---- *)
FUNCTION_BLOCK HTML_DECODE

	VAR_INPUT
		IN :	oscat_STRING250;
	END_VAR

	VAR_OUTPUT
		HTML_DECODE :	oscat_STRING250;
	END_VAR

	VAR
		pos :	INT;
		end :	INT;
		tmp :	oscat_STRING10;
		code :	BYTE;
		size :	INT;
		CHR_TO_STRING :	CHR_TO_STRING;
		CHARCODE :	CHARCODE;
		HEX_TO_DWORD :	HEX_TO_DWORD;
		FINDP :	FINDP;
	END_VAR

	HTML_DECODE := IN;

	pos := FIND(HTML_DECODE, '&');
	WHILE pos > 0 DO
		tmp := MID(HTML_DECODE, 2, pos + 1);
		IF EQ_STRING(tmp,'#x') OR EQ_STRING(tmp,'#X') THEN

			IF pos+13 > LEN(HTML_DECODE) THEN
			size := LEN(HTML_DECODE) - pos - 2;
			ELSE
			size := 10;
			END_IF;

			tmp := MID(HTML_DECODE, size, pos + 3);
			end := FIND(tmp, ';');
			HEX_TO_DWORD(Hex:=LEFT(tmp, end - 1));
			CODE := DWORD_TO_BYTE(HEX_TO_DWORD.HEX_TO_DWORD);
			CHR_TO_STRING(C:=CODE);
			HTML_DECODE := REPLACE(HTML_DECODE, CHR_TO_STRING.CHR_TO_STRING, end + 3, pos);
		ELSE
			tmp := LEFT(tmp,1);
			IF EQ_STRING(tmp,'#') THEN

				IF pos+12 > LEN(HTML_DECODE) THEN
					size := LEN(HTML_DECODE) - pos - 1;
				ELSE
					size := 10;
				END_IF;

				tmp := MID(HTML_DECODE, size, pos + 2);
				end := FIND(tmp, ';');
				tmp := LEFT(tmp, end - 1);
				CODE := INT_TO_BYTE(STRING_TO_INT(tmp));
				CHR_TO_STRING(C:=CODE);
				HTML_DECODE := REPLACE(HTML_DECODE, CHR_TO_STRING.CHR_TO_STRING, end + 2, pos);
			ELSE
				IF pos+11 > LEN(HTML_DECODE) THEN
					size := LEN(HTML_DECODE) - pos ;
				ELSE
					size := 10;
				END_IF;

				tmp := MID(HTML_DECODE, size, pos + 1);
				end := FIND(tmp, ';');
				CHARCODE(STR:=LEFT(tmp, end - 1));
				CODE := CHARCODE.CHARCODE;
				CHR_TO_STRING(C:=CODE);
				HTML_DECODE := REPLACE(HTML_DECODE, CHR_TO_STRING.CHR_TO_STRING, end + 1, pos);
			END_IF;
		END_IF;
		FINDP(str:=HTML_DECODE,src:='&',pos:=pos + 1);
		pos := FINDP.FINDP;
	END_WHILE;

END_FUNCTION_BLOCK

(* ---- HTML_ENCODE.ST ---- *)
FUNCTION_BLOCK HTML_ENCODE

	VAR_INPUT
		IN :	oscat_STRING250;
		M :	BOOL;
	END_VAR

	VAR_OUTPUT
		HTML_ENCODE :	oscat_STRING250;
	END_VAR

	VAR
		pt_out :	oscat_aB1_255;
		pos_in :	INT;
		pos_out :	INT;
		stop :	INT;
		B :	INT;
		tmp :	oscat_STRING10;
		i :	INT;
		BUF_TO_STRING :	BUF_TO_STRING;
		CHARNAME :	CHARNAME;
		CODE :	CODE;
	END_VAR

	pos_in := 1;
	stop := LEN(in);
	FOR pos_out := 1 TO 250 DO
		IF pos_in > stop THEN EXIT; END_IF;
		B := GET_CHAR(IN,pos_in);
		CASE B OF
			34:
				IF pos_out > 244 THEN EXIT; END_IF;
				pt_out[pos_out] := BYTE#38;
				pos_out := pos_out + 1;
				pt_out[pos_out] := BYTE#113;
				pos_out := pos_out + 1;
				pt_out[pos_out] := BYTE#117;
				pos_out := pos_out + 1;
				pt_out[pos_out] := BYTE#111;
				pos_out := pos_out + 1;
				pt_out[pos_out] := BYTE#116;
				pos_out := pos_out + 1;
				pt_out[pos_out] := BYTE#59;
			38:
				IF pos_out > 245 THEN EXIT; END_IF;
				pt_out[pos_out] := BYTE#38;
				pos_out := pos_out + 1;
				pt_out[pos_out] := BYTE#97;
				pos_out := pos_out + 1;
				pt_out[pos_out] := BYTE#109;
				pos_out := pos_out + 1;
				pt_out[pos_out] := BYTE#112;
				pos_out := pos_out + 1;
				pt_out[pos_out] := BYTE#59;
			60:
				IF pos_out > 246 THEN EXIT; END_IF;
				pt_out[pos_out] := BYTE#38;
				pos_out := pos_out + 1;
				pt_out[pos_out] := BYTE#108;
				pos_out := pos_out + 1;
				pt_out[pos_out] := BYTE#116;
				pos_out := pos_out + 1;
				pt_out[pos_out] := BYTE#59;
			62:
				IF pos_out > 246 THEN EXIT; END_IF;
				pt_out[pos_out] := BYTE#38;
				pos_out := pos_out + 1;
				pt_out[pos_out] := BYTE#103;
				pos_out := pos_out + 1;
				pt_out[pos_out] := BYTE#116;
				pos_out := pos_out + 1;
				pt_out[pos_out] := BYTE#59;
		ELSE
			IF M AND B > 127 THEN
				CHARNAME(C:=INT_TO_BYTE(B));
				tmp := CHARNAME.CHARNAME;
				IF pos_out + LEN(tmp) + 2 <= 250 THEN
					pt_out[pos_out] := BYTE#38;
					pos_out := pos_out + 1;
					FOR i := 1 TO LEN(tmp) DO
						CODE(STR:=tmp,POS:=i);
						pt_out[pos_out] := CODE.CODE;
						pos_out := pos_out + 1;
					END_FOR;
					pt_out[pos_out] := BYTE#59;
				END_IF;
			ELSE
			pt_out[pos_out] := INT_TO_BYTE(B);
			END_IF;
		END_CASE;
		pos_in := pos_in + 1;
	END_FOR;

	pos_out := pos_out - 1;

	FOR pos_in := 0 TO 1 DO
	BUF_TO_STRING.REQ        := pos_in>0;
	BUF_TO_STRING.BUF_FORMAT := TRUE;
	BUF_TO_STRING.BUF_OFFS   := DINT#0;
	BUF_TO_STRING.BUF_CNT    := INT_TO_DINT(pos_out);
	BUF_TO_STRING.BUFFER     := pt_out;
	BUF_TO_STRING.DST        := HTML_ENCODE;
	BUF_TO_STRING();
	pt_out  := BUF_TO_STRING.BUFFER;
	HTML_ENCODE := BUF_TO_STRING.DST;
	END_FOR;

END_FUNCTION_BLOCK

(* ---- HYST.ST ---- *)
FUNCTION_BLOCK HYST_Block

	VAR_INPUT
		IN :	REAL;
		_ON :	REAL;
		OFF :	REAL;
	END_VAR

	VAR_OUTPUT
		Q :	BOOL;
		WIN :	BOOL;
	END_VAR

	IF _ON >= OFF THEN
		IF IN < OFF THEN
			Q := FALSE;
			WIN := FALSE;
		ELSIF  IN > _ON THEN
			Q := TRUE;
			WIN := FALSE;
		ELSE
			WIN := TRUE;
		END_IF;
	ELSE
		IF IN > OFF THEN
			Q := FALSE;
			WIN := FALSE;
		ELSIF  IN < _ON THEN
			Q := TRUE;
			WIN := FALSE;
		ELSE
			WIN := TRUE;
		END_IF;
	END_IF;

END_FUNCTION_BLOCK

PROGRAM program0
	VAR
		IN :	REAL;
		_ON :	REAL;
		OFF :	REAL;
		Q :	BOOL;
		WIN :	BOOL;
		func_block : HYST_Block;
	END_VAR
	func_block.IN := IN;
	func_block._ON := _ON;
	func_block.OFF := OFF ;
	func_block();
	Q  := func_block.Q;
	WIN  := func_block.WIN;
END_PROGRAM

CONFIGURATION Config0
	RESOURCE Res0 ON PLC
		TASK task0(INTERVAL := T#20ms,PRIORITY := 0);
		PROGRAM instance0 WITH task0 : program0;
	END_RESOURCE
END_CONFIGURATION

(* ---- HYST_1.ST ---- *)
FUNCTION_BLOCK HYST_1_Block

	VAR_INPUT
		IN :	REAL;
		HIGH :	REAL;
		LOW :	REAL;
	END_VAR

	VAR_OUTPUT
		Q :	BOOL;
		WIN :	BOOL;
	END_VAR

	IF in < low THEN
		Q := FALSE;
		win := FALSE;
	ELSIF in > high THEN
		Q := TRUE;
		win := FALSE;
	ELSE
		win := TRUE;
	END_IF;

END_FUNCTION_BLOCK

PROGRAM program0
	VAR
		IN :	REAL;
		HIGH :	REAL;
		LOW :	REAL;
		Q :	BOOL;
		WIN :	BOOL;
		func_block : HYST_1_Block;
	END_VAR
	func_block.IN := IN;
	func_block.HIGH := HIGH;
	func_block.LOW := LOW;
	func_block();
	Q  := func_block.Q;
	WIN  := func_block.WIN;
END_PROGRAM

CONFIGURATION Config0
	RESOURCE Res0 ON PLC
		TASK task0(INTERVAL := T#20ms,PRIORITY := 0);
		PROGRAM instance0 WITH task0 : program0;
	END_RESOURCE
END_CONFIGURATION

(* ---- HYST_2.ST ---- *)
FUNCTION_BLOCK HYST_2_Block

	VAR_INPUT
		IN :	REAL;
		VAL :	REAL;
		HYS :	REAL;
	END_VAR

	VAR_OUTPUT
		Q :	BOOL;
		WIN :	BOOL;
	END_VAR

	VAR
		tmp :	REAL;
	END_VAR

	tmp := val - hys * 0.5;
	IF in < tmp THEN
		Q := FALSE;
		win := FALSE;
	ELSIF in > tmp + hys THEN
		Q := TRUE;
		win := FALSE;
	ELSE
		win := TRUE;
	END_IF;

END_FUNCTION_BLOCK

PROGRAM program0
	VAR
		IN :	REAL;
		VAL :	REAL;
		HYS :	REAL;
		Q :	BOOL;
		WIN :	BOOL;
		func_block : HYST_2_Block;
	END_VAR
	func_block.IN := IN;
	func_block.VAL := VAL;
	func_block.HYS := HYS;
	func_block();
	Q  := func_block.Q;
	WIN  := func_block.WIN;
END_PROGRAM

CONFIGURATION Config0
	RESOURCE Res0 ON PLC
		TASK task0(INTERVAL := T#20ms,PRIORITY := 0);
		PROGRAM instance0 WITH task0 : program0;
	END_RESOURCE
END_CONFIGURATION

(* ---- HYST_3.ST ---- *)
FUNCTION_BLOCK HYST_3_Block

	VAR_INPUT
		IN :	REAL;
		HYST :	REAL;
		VAL1 :	REAL;
		VAL2 :	REAL;
	END_VAR

	VAR_OUTPUT
		Q1 :	BOOL;
		Q2 :	BOOL;
	END_VAR

	VAR
		X :	REAL;
	END_VAR

	X := hyst * 0.5;
	IF in < val1 - X THEN
		q1 := TRUE;
	ELSIF in > val1 + X THEN
		q1 := FALSE;
	END_IF;
	IF in < val2 - X THEN
		q2 := FALSE;
	ELSIF in > val2 + X THEN
		q2 := TRUE;
	END_IF;

END_FUNCTION_BLOCK

PROGRAM program0
	VAR
		IN :	REAL;
		HYST :	REAL;
		VAL1 :	REAL;
		VAL2 :	REAL;
		Q1 :	BOOL;
		Q2 :	BOOL;
		func_block : HYST_3_Block;
	END_VAR
	func_block.IN := IN;
	func_block.HYST := HYST;
	func_block.VAL1 := VAL1;
	func_block.VAL2 := VAL2;
	func_block();
	Q1  := func_block.Q1;
	Q2  := func_block.Q2;
END_PROGRAM

CONFIGURATION Config0
	RESOURCE Res0 ON PLC
		TASK task0(INTERVAL := T#20ms,PRIORITY := 0);
		PROGRAM instance0 WITH task0 : program0;
	END_RESOURCE
END_CONFIGURATION

(* ---- INC_DEC.ST ---- *)
FUNCTION_BLOCK INC_DEC_Block

	VAR_INPUT
		CHA :	BOOL;
		CHB :	BOOL;
		RST :	BOOL := 0;
	END_VAR

	VAR_OUTPUT
		DIR :	BOOL;
		CNT :	INT;
	END_VAR

	VAR
		edgea :	BOOL := 0;
		clk :	BOOL;
		clka :	BOOL;
		clkb :	BOOL;
		edgeb :	BOOL;
		axb :	BOOL;
	END_VAR

	axb := cha XOR chb;

	clka := cha XOR edgea;
	edgea := cha;

	clkb := chb XOR edgeb;
	edgeb := chb;

	clk := clka OR clkb;

	IF axb AND clka THEN dir := TRUE; END_IF;
	IF axb AND clkb THEN dir := FALSE; END_IF;

	IF clk AND dir THEN cnt := cnt + 1; END_IF;
	IF clk AND NOT dir THEN cnt := cnt -1; END_IF;

	IF rst THEN cnt := 0; END_IF;

END_FUNCTION_BLOCK

PROGRAM program0

	VAR
		CHA :	BOOL;
		CHB :	BOOL;
		RST :	BOOL := 0;

		DIR :	BOOL;
		CNT :	INT;
		func_block : INC_DEC_Block;
	END_VAR
	func_block.CHA := CHA;
	func_block.CHB := CHB;
	func_block.RST := RST;
	func_block();
	DIR := func_block.DIR;
	CNT := func_block.CNT;

END_PROGRAM

CONFIGURATION Config0

	RESOURCE Res0 ON PLC
		TASK task0(INTERVAL := T#20ms,PRIORITY := 0);
		PROGRAM instance0 WITH task0 : program0;
	END_RESOURCE

END_CONFIGURATION

(* ---- INSERT250.ST ---- *)
TYPE
	oscat_STRING250             : STRING;
END_TYPE

FUNCTION_BLOCK _INSERT250
    VAR_INPUT
        IN1 :	oscat_STRING250;
        IN2 :	oscat_STRING250;
        P :	INT;
    END_VAR
    VAR_OUTPUT
        _INSERT :	oscat_STRING250;
    END_VAR
    VAR
        size :	INT;
    END_VAR

    size := LEN(IN1);
    IF size + LEN(IN2) <= 250 THEN
        P := LIMIT(0,P,size);
        IF P = 0 THEN
            _INSERT := CONCAT(IN2,IN1);
        ELSE
            _INSERT := INSERT(IN1, IN2, P);
        END_IF;
    END_IF;

END_FUNCTION_BLOCK

PROGRAM program0
	VAR
	    LocalVar1 : oscat_STRING250;
        LocalVar2 : oscat_STRING250;
        LocalVar3 : INT;
		LocalOUT  : oscat_STRING250;
		func_block : _INSERT250;
  	END_VAR
	func_block.IN1 := LocalVar1;
    func_block.IN2 := LocalVar2;
    func_block.P := LocalVar3;
	func_block();
	LocalOUT := func_block._INSERT;
END_PROGRAM

CONFIGURATION Config0
  	RESOURCE Res0 ON PLC
    	TASK task0(INTERVAL := T#20ms,PRIORITY := 0);
    	PROGRAM instance0 WITH task0 : program0;
  	END_RESOURCE
END_CONFIGURATION

(* ---- INTEGRATE.ST ---- *)
FUNCTION_BLOCK T_PLC_MS_block
	VAR_OUTPUT
		T_PLC_MS :	UDINT;
	END_VAR

	VAR_EXTERNAL
		PLC_TICKS_PER_SEC :	INT;
		PLC_SYS_TICK_CNT :	DINT;
	END_VAR

	VAR
		debug :	BOOL;(*Debug-Mode ON / OFF*)
		N :	INT;(*Debug-Faktor*)
		Offset :	UDINT;(*Debug-Offset*)
		temp :	DWORD := DWORD#1;(*Debug-Offset*)
		mode :	BOOL;(*modus*)
		faktor :	UDINT;(*Systemtakt-Faktor*)
		init :	BOOL;
		v_plc_ticks_per_sec :	UDINT;
		base :	UDINT := UDINT#1000;
	END_VAR

	IF init = FALSE THEN
		v_plc_ticks_per_sec := INT_TO_UDINT(PLC_TICKS_PER_SEC);
		IF v_plc_ticks_per_sec = UDINT#1024 THEN
			faktor := UDINT#1;
			mode := FALSE;
		ELSIF v_plc_ticks_per_sec > UDINT#0 THEN
			IF v_plc_ticks_per_sec <= base THEN
				faktor := base / v_plc_ticks_per_sec;
				mode := FALSE;
			ELSE
				faktor := v_plc_ticks_per_sec / base;
				mode := TRUE;
			END_IF;
		ELSE
			faktor := UDINT#1;
		END_IF;
		init := TRUE;
	END_IF;

	IF mode THEN
		T_PLC_MS := DINT_TO_UDINT(PLC_SYS_TICK_CNT) / faktor;
	ELSE
		T_PLC_MS := DINT_TO_UDINT(PLC_SYS_TICK_CNT) * faktor;
	END_IF;

	IF debug THEN
		T_PLC_MS := (DWORD_TO_UDINT(SHL(UDINT_TO_DWORD(T_PLC_MS),N) OR SHL(temp,N)) - UDINT#1) + Offset;
	END_IF;
END_FUNCTION_BLOCK

FUNCTION_BLOCK INTEGRATE

	VAR_INPUT
		E :	BOOL := TRUE;
		X :	REAL;
		K :	REAL := 1.0;
	END_VAR

	VAR_IN_OUT
		Y :	REAL;
	END_VAR

	VAR
		X_last :	REAL;
		init :	BOOL;
		T_PLC_MS :	T_PLC_MS_block;
		last :	UDINT;
		tx :	UDINT;
	END_VAR

	T_PLC_MS();
	tx:= T_PLC_MS.T_PLC_MS;

	IF NOT init THEN
		init := TRUE;
		X_last := X;
	ELSIF E THEN
		Y := (X + X_LAST) * 0.5E-3 * UDINT_TO_REAL(tx-last) * K + Y;
		X_last := X;
	END_IF;
	last := tx;

END_FUNCTION_BLOCK

PROGRAM program0
  VAR
	E :	BOOL := TRUE;
	X :	REAL;
	K :	REAL := 1.0;

	Y :	REAL;

	func_block : INTEGRATE;
  END_VAR
	func_block.E:=E;
	func_block.X:=X;
	func_block.K:=K;
	func_block.Y:=Y;
	func_block();
	Y:= func_block.Y;
END_PROGRAM

CONFIGURATION Config0
	VAR_GLOBAL
		PLC_TICKS_PER_SEC :	INT;
		PLC_SYS_TICK_CNT :	DINT;
	END_VAR
	RESOURCE Res0 ON PLC
		TASK task0(INTERVAL := T#20ms,PRIORITY := 0);
		PROGRAM instance0 WITH task0 : program0;
	END_RESOURCE
END_CONFIGURATION

(* ---- INTERLOCK.ST ---- *)
FUNCTION_BLOCK INTERLOCK_Block

	VAR_INPUT
		I1 :	BOOL;
		I2 :	BOOL;
		TL :	TIME;
	END_VAR

	VAR_OUTPUT
		Q1 :	BOOL;
		Q2 :	BOOL;
	END_VAR

	VAR
		T1 :	TOF;
		T2 :	TOF;
	END_VAR

	T1(IN := I1, PT := TL);
	T2(IN := I2, PT := TL);

	Q1 := I1 AND NOT t2.Q;
	Q2 := I2 AND NOT t1.Q;

END_FUNCTION_BLOCK

PROGRAM program0
	VAR
		I1 :	BOOL;
		I2 :	BOOL;
		TL :	TIME;
		Q1 :	BOOL;
		Q2 :	BOOL;
		func_block : INTERLOCK_Block;
  	END_VAR
	func_block.I1  :=I1;
	func_block.I2  :=I2;
	func_block.TL  :=TL;
	func_block();
	Q1 := func_block.Q1;
	Q2 := func_block.Q2;
END_PROGRAM

CONFIGURATION Config0
	RESOURCE Res0 ON PLC
		TASK task0(INTERVAL := T#20ms,PRIORITY := 0);
		PROGRAM instance0 WITH task0 : program0;
	END_RESOURCE
END_CONFIGURATION

(* ---- INTERLOCK_4.ST ---- *)
FUNCTION BIT_LOAD_B:BYTE
	VAR_INPUT
		IN :	BYTE;
		VAL :	BOOL;
		POS :	INT;
	END_VAR

	IF VAL THEN
		BIT_LOAD_B := in OR SHL(BYTE#1,pos);
	ELSE
		BIT_LOAD_B := in AND (NOT SHL(BYTE#1,pos));
	END_IF;
END_FUNCTION

FUNCTION_BLOCK INTERLOCK_4_Block

	VAR_INPUT
		I0 :	BOOL;
		I1 :	BOOL;
		I2 :	BOOL;
		I3 :	BOOL;
		E :	BOOL;
		MODE :	INT;
	END_VAR

	VAR_OUTPUT
		OUT :	BYTE;
		_TP :	BOOL;
	END_VAR

	VAR
		in :	BYTE;
		last :	BYTE;
		old :	BYTE;
		lmode :	INT;
	END_VAR

	IF E THEN
	(* reset all vars when there is a mode change on thy fly *)
		IF mode <> lmode THEN
			out := BYTE#0;
			last := BYTE#0;
			old := BYTE#0;
			lmode := mode;
		END_IF;
		(* load inputs into in *)
		in:=BIT_LOAD_B(in,I0,0); (* in.0 *)
		in:=BIT_LOAD_B(in,I1,1); (* in.1 *)
		in:=BIT_LOAD_B(in,I2,2); (* in.2 *)
		in:=BIT_LOAD_B(in,I3,3); (* in.3 *)
		(* only execute when there is any change *)
		IF in <> last THEN
			(* only execute when inputs have chages state *)
			CASE mode OF
				0:	(* output directly display inputs as bits in byte out *)
					out := in;

				1:	(* the input with the highest number will be acepted *)
					IF    (in AND BYTE#2#00001000) > BYTE#0 (* in.3 *) THEN out := BYTE#8;
					ELSIF (in AND BYTE#2#00000100) > BYTE#0 (* in.2 *) THEN out := BYTE#4;
					ELSIF (in AND BYTE#2#00000010) > BYTE#0 (* in.1 *) THEN out := BYTE#2;
					ELSE out := in;
					END_IF;

				2:	(* input last pressed will be displayed only *)
					last := ((in XOR last) AND in);
					IF    (last AND BYTE#2#00001000) > BYTE#0 (* last.3 *) THEN out := BYTE#8;
					ELSIF (last AND BYTE#2#00000100) > BYTE#0 (* last.2 *) THEN out := BYTE#4;
					ELSIF (last AND BYTE#2#00000010) > BYTE#0 (* last.1 *) THEN out := BYTE#2;
					ELSE out := last;
					END_IF;

				3:	(* any input active will disable all other inputs *)
					IF (out AND in) = BYTE#0 THEN
						IF    (in AND BYTE#2#00001000) > BYTE#0 (* in.3 *) THEN out := BYTE#8;
						ELSIF (in AND BYTE#2#00000100) > BYTE#0 (* in.2 *) THEN out := BYTE#4;
						ELSIF (in AND BYTE#2#00000010) > BYTE#0 (* in.1 *) THEN out := BYTE#2;
						ELSE out := in;
						END_IF;
					END_IF;

			END_CASE;
			last := in;
		END_IF;
		_tp := out <> old;
		old := out;
	ELSE
		out := BYTE#0;
		last := BYTE#0;
		old := BYTE#0;
		lmode := 0;
		_tp := FALSE;
	END_IF;

END_FUNCTION_BLOCK

PROGRAM program0

	VAR
		I0 :	BOOL;
		I1 :	BOOL;
		I2 :	BOOL;
		I3 :	BOOL;
		E :	BOOL;
		MODE :	INT;
		OUT :	BYTE;
		_TP :	BOOL;
		func_block : INTERLOCK_4_Block;
	END_VAR
	func_block.I0 := I0;
	func_block.I1 := I1;
	func_block.I2 := I2;
	func_block.I3 := I3;
	func_block.E := E;
	func_block.MODE := MODE;
	func_block();
	OUT := func_block.OUT;
	_TP := func_block._TP;

END_PROGRAM

CONFIGURATION Config0

	RESOURCE Res0 ON PLC
		TASK task0(INTERVAL := T#20ms,PRIORITY := 0);
		PROGRAM instance0 WITH task0 : program0;
	END_RESOURCE

END_CONFIGURATION

(* ---- IP2GEO.ST ---- *)
FUNCTION_BLOCK IP2GEO

  VAR_IN_OUT
    IP_C :	oscat_IP_C;
    S_BUF :	oscat_NETWORK_BUFFER;
    R_BUF :	oscat_NETWORK_BUFFER;
    GEO :	oscat_IP2GEO_DATA;
  END_VAR

  VAR_INPUT
    IP :	DWORD;
    ACTIVATE :	BOOL;
  END_VAR

  VAR_OUTPUT
    BUSY :	BOOL;
    DONE :	BOOL;
    ERROR_C :	DWORD;
    ERROR_T :	BYTE;
  END_VAR

  VAR
    CTRL :	oscat_XML_CONTROL;
    XML_READER :	XML_READER;
    URL_DATA :	oscat_url;
    DNS_CLIENT :	DNS_CLIENT;
    STRING_TO_URL :	STRING_TO_URL;
    HTTP_GET :	HTTP_GET;
    FLOAT_TO_REAL :	FLOAT_TO_REAL;
    last_state :	BOOL;
    value_int :	INT;
    value_real :	REAL;
    v_real :	REAL;
    state :	INT;
    IP4_TO_STRING :	IP4_TO_STRING;
    IP4_DECODE :	IP4_DECODE;
    CHK_REAL :	CHK_REAL;
  END_VAR

  CASE state OF

  00:
    IF ACTIVATE AND NOT last_state THEN
      state := 20;
    DONE := FALSE;
    BUSY := TRUE;
    ERROR_C := DWORD#0;
    ERROR_T := BYTE#0;
    END_IF;

  20:
    STRING_TO_URL.STR:='http://ipinfodb.com/ip_query.php?timezone=true&IP=';
    STRING_TO_URL.DEFAULT_PROTOCOL:='';
    STRING_TO_URL.DEFAULT_PATH:='';
    STRING_TO_URL();
    URL_DATA:=STRING_TO_URL.STRING_TO_URL;

    IF IP > DWORD#0 THEN
      IP4_TO_STRING(IP4:=IP);
      URL_DATA.QUERY := CONCAT(URL_DATA.QUERY,IP4_TO_STRING.IP4_TO_STRING);
    END_IF;

    state := 40;

  40:
    IF DNS_CLIENT.DONE THEN
      state := 60;
    ELSIF (DNS_CLIENT.ERROR > DWORD#00) THEN
      ERROR_C := DNS_CLIENT.ERROR;
    ERROR_T := BYTE#01;
      state   := 100;
    END_IF;

  60:
    IF HTTP_GET.DONE THEN
      state := 80;
      CTRL.START_POS := HTTP_GET.BODY_START;
      CTRL.STOP_POS  := HTTP_GET.BODY_STOP;
      CTRL.COMMAND   := WORD#2#10000000_00011000;
    CTRL.WATCHDOG  := T#1ms;

    ELSIF (HTTP_GET.ERROR > DWORD#00) THEN
      ERROR_C := HTTP_GET.ERROR;
      ERROR_T := BYTE#02;
      state   := 100;
    END_IF;

  80:
    XML_READER.CTRL := CTRL;
    XML_READER.BUF  := R_BUF.BUFFER;
    XML_READER();
    CTRL         := XML_READER.CTRL;
    R_BUF.BUFFER := XML_READER.BUF;

    IF CTRL.TYP < 98 THEN
      value_int := 0;
      value_real := 0.0;
      IF LEN(CTRL.VALUE) <= 20 THEN
            FLOAT_TO_REAL(FLT:=CTRL.VALUE);
        v_real :=FLOAT_TO_REAL.FLOAT_TO_REAL;
        CHK_REAL(X:= v_real);
        IF CHK_REAL.CHK_REAL = BYTE#0 THEN
          value_real := v_real;
          value_int := REAL_TO_INT(value_real);
        END_IF;
      END_IF;

      CASE UINT_TO_INT(CTRL.COUNT) OF

        07: IP4_DECODE(STR:=CTRL.VALUE);
            GEO.IP4 := IP4_DECODE.IP4_DECODE;
      10: GEO.STATE := EQ_STRING('OK',CTRL.VALUE);
      13: GEO.COUNTRY_CODE := CTRL.VALUE;
      16: GEO.COUNTRY_NAME := CTRL.VALUE;
      19: GEO.REGION_CODE := CTRL.VALUE;
      22: GEO.REGION_NAME := CTRL.VALUE;
      25: GEO.CITY := CTRL.VALUE;
      31: GEO.GEO_LATITUDE := value_real;
      34: GEO.GEO_LONGITUDE := value_real;
      37: GEO.TIME_ZONE_NAME := CTRL.VALUE;
      40: GEO.GMT_OFFSET := value_int;
      43: GEO.IS_DST := value_int > 0;
      END_CASE;

    ELSIF CTRL.TYP = 99 THEN
      DONE  := TRUE;
      state := 100;
    END_IF;

  100:
    IF (NOT HTTP_GET.DONE) THEN
      state := 0;
      BUSY  := FALSE;
      DONE := ERROR_T = BYTE#0;
    END_IF;

  END_CASE;

  DNS_CLIENT.IP_C     := IP_C;
  DNS_CLIENT.S_BUF    := S_BUF;
  DNS_CLIENT.R_BUF    := R_BUF;
  DNS_CLIENT.DOMAIN   := URL_DATA.DOMAIN;
  DNS_CLIENT.IP4_DNS  := DWORD#00;
  DNS_CLIENT.ACTIVATE := state=40;
  DNS_CLIENT();
  IP_C  := DNS_CLIENT.IP_C;
  S_BUF := DNS_CLIENT.S_BUF;
  R_BUF := DNS_CLIENT.R_BUF;

  HTTP_GET.IP_C        := IP_C;
  HTTP_GET.S_BUF       := S_BUF;
  HTTP_GET.R_BUF       := R_BUF;
  HTTP_GET.IP4         := DNS_CLIENT.IP4;
  HTTP_GET.GET         := state=60;
  HTTP_GET.MODE        := BYTE#2;
  HTTP_GET.UNLOCK_BUF  := state=100;
  HTTP_GET.URL_DATA    := URL_DATA;
  HTTP_GET();
  IP_C     := HTTP_GET.IP_C;
  S_BUF    := HTTP_GET.S_BUF;
  R_BUF    := HTTP_GET.R_BUF;
  URL_DATA := HTTP_GET.URL_DATA;

  last_state := ACTIVATE;

END_FUNCTION_BLOCK

(* ---- IP4_DECODE.ST ---- *)
TYPE
  oscat_STRING80             : STRING;
END_TYPE

FUNCTION_BLOCK IP4_DECODE_Block

	VAR_INPUT
		STR :	oscat_STRING80;
	END_VAR

	VAR_OUTPUT
		IP4_DECODE :	DWORD;
	END_VAR

	VAR
		pos :	INT;
		IS_NUM :	IS_NUM;
	END_VAR

	IP4_DECODE := DWORD#0;
	pos := FIND(str, '.');
	WHILE pos > 0 DO
		IP4_DECODE := SHL(IP4_DECODE,8);
		IF POS > 1 AND POS <= 4 THEN
			IS_NUM(STR:=LEFT(str,pos - 1));
			IF IS_NUM.IS_NUM THEN
				IP4_DECODE := IP4_DECODE OR STRING_TO_DWORD(IS_NUM.STR);
			END_IF;
		END_IF;
		str := DELETE(str, pos, 1);
		pos := FIND(str, '.');
	END_WHILE;

	IP4_DECODE := SHL(IP4_DECODE,8);
	IS_NUM(STR:=str);
	IF IS_NUM.IS_NUM THEN
	IP4_DECODE := IP4_DECODE OR STRING_TO_DWORD(str);
	END_IF;

END_FUNCTION_BLOCK

PROGRAM program0
	VAR
		STR :	oscat_STRING80;
		IP4_DECODE :	DWORD;

		func_block : IP4_DECODE_Block;
	END_VAR
	func_block.STR := STR;

	func_block();
	IP4_DECODE  := func_block.IP4_DECODE;
END_PROGRAM

CONFIGURATION Config0

  	RESOURCE Res0 ON PLC
    	TASK task0(INTERVAL := T#20ms,PRIORITY := 0);
    	PROGRAM instance0 WITH task0 : program0;
  	END_RESOURCE

END_CONFIGURATION

(* ---- IP4_TO_STRING.ST ---- *)
TYPE
  oscat_STRING10             : STRING;
END_TYPE

FUNCTION _BYTE_TO_INT:INT
	VAR_INPUT
		IN :	BYTE;
	END_VAR

	_BYTE_TO_INT := USINT_TO_INT(BYTE_TO_USINT(IN));
END_FUNCTION

FUNCTION BYTE_OF_DWORD:BYTE
	VAR_INPUT
		IN :	DWORD;
		N :	BYTE;
	END_VAR
	BYTE_OF_DWORD := DWORD_TO_BYTE(SHR(in,_BYTE_TO_INT(SHL(n,3))));
END_FUNCTION

FUNCTION_BLOCK IP4_TO_STRING_Block

	VAR_INPUT
		IP4 :	DWORD;
	END_VAR

	VAR_OUTPUT
		IP4_TO_STRING :	STRING;
	END_VAR

	VAR
		s1 :	oscat_string10;
		s2 :	oscat_string10;
	END_VAR

	s1 := CONCAT(BYTE_TO_STRING(BYTE_OF_DWORD(IP4,BYTE#1)),BYTE_TO_STRING(BYTE_OF_DWORD(IP4,BYTE#0)));
	s2 := CONCAT(BYTE_TO_STRING(BYTE_OF_DWORD(IP4,BYTE#3)),BYTE_TO_STRING(BYTE_OF_DWORD(IP4,BYTE#2)));
	IP4_TO_STRING := CONCAT(s2,s1);

END_FUNCTION_BLOCK

PROGRAM program0
	VAR
		IP4 :	DWORD;
		IP4_TO_STRING :	STRING;

		func_block : IP4_TO_STRING_Block;
	END_VAR
	func_block.IP4 := IP4;

	func_block();
	IP4_TO_STRING  := func_block.IP4_TO_STRING;
END_PROGRAM

CONFIGURATION Config0

  	RESOURCE Res0 ON PLC
    	TASK task0(INTERVAL := T#20ms,PRIORITY := 0);
    	PROGRAM instance0 WITH task0 : program0;
  	END_RESOURCE

END_CONFIGURATION

(* ---- IP_CONTROL.ST ---- *)
FUNCTION_BLOCK IP_CONTROL_Block

  VAR
    T_PLC_MS :	T_PLC_MS;
    IP4_TO_STRING :	IP4_TO_STRING;
    FB_IP_CONNECT :	IP_CONNECT;
    FB_IP_URCV :	IP_URCV;
    FB_IP_USEND :	IP_USEND;
  END_VAR

  VAR_INPUT
    IP :	DWORD;
    PORT :	WORD;
    TIME_OUT :	TIME;
  END_VAR

  VAR_IN_OUT
    IP_C :	oscat_IP_C;
    S_BUF :	oscat_NETWORK_BUFFER;
    R_BUF :	oscat_NETWORK_BUFFER;
  END_VAR

  VAR
    C_TIME :	UDINT;
    S_TIME :	UDINT;
    R_TIME :	UDINT;
    C_ENABLE :	BOOL;
    C_IP :	DWORD;
    C_PORT :	WORD;
    C_MODE :	BYTE;
    C_ERROR :	BOOL;
    C_STATUS :	INT;
    C_ID :	INT;
    C_RECONNECT :	BOOL;
    C_RECONNECT_COUNT :	INT;
    S_BUF_I :	oscat_NETWORK_BUFFER_SHORT;
    S_TOTAL :	INT;
    S_CUR_POS :	INT;
    S_CUR_SIZE :	INT;
    S_MAX_SIZE :	INT := 1408;
    S_START :	BOOL;
    S_REQ :	BOOL;
    S_DONE :	BOOL;
    S_ERROR :	BOOL;
    S_STATUS :	INT;
    R_NDR :	BOOL;
    R_ERROR :	BOOL;
    R_STATUS :	INT;
    R_BUF_I :	oscat_NETWORK_BUFFER_SHORT;
    R_COUNT :	INT;
    R_OFFSET :	INT;
    R_E_MAX_SIZE :	INT := 4096;
    NEW_CONNECTION :	BOOL;
    C_ENABLE_OLD :	BOOL;
    C_READY :	BOOL;
    C_READY_OLD :	BOOL;
    DELAY_STOP :	UDINT;
    DELAY :	UDINT;
    DELAY_VALUE :	UDINT;
    C :	INT;
    C2 :	INT;
    C3 :	INT;
    CS :	STRING;
    TX :	UDINT;
    ERROR_TIME :	UDINT;
    S_ACTIVE :	BOOL;
    ERROR_CON :	BYTE;
    ERROR_SND :	BYTE;
    ERROR_RCV :	BYTE;
  END_VAR

  T_PLC_MS();
  TX := T_PLC_MS.T_PLC_MS;

  IF (TX - DELAY < DELAY_VALUE) THEN
    IF IP_C.C_STATE <> BYTE#1 AND IP_C.C_STATE <> BYTE#254 THEN
    RETURN;
    END_IF;
  END_IF;
  DELAY := TX;

  IF C_ENABLE AND DELAY_VALUE > UDINT#00 THEN
    IF (TX - DELAY_STOP > UDINT#1000) THEN
      DELAY_VALUE := UDINT#00;
    END_IF;
  ELSE
    DELAY_STOP := TX;
  END_IF;

  IF IP_C.C_PORT = WORD#00 THEN
    IP_C.C_PORT := PORT;
  END_IF;
  IF IP_C.C_IP=DWORD#00 AND IP_C.C_MODE<BYTE#4 THEN
    IP_C.C_IP := IP;
  END_IF;

  NEW_CONNECTION := C_IP <> IP_C.C_IP OR C_MODE <> IP_C.C_MODE OR C_PORT <> IP_C.C_PORT;

  IF IP_C.C_ENABLE AND NOT C_READY AND NEW_CONNECTION THEN

    C_IP   := IP_C.C_IP;
    C_MODE := IP_C.C_MODE;
    C_PORT := IP_C.C_PORT;

    CS := SEL_STRING((C_MODE AND BYTE#1) = BYTE#1,'','/UDP');
    CS := CONCAT(CS,SEL_STRING(C_MODE<BYTE#2,' /PASSIVE',' /ACTIVE'));
    CS := CONCAT(CS,' /PORT=');
    CS := CONCAT(CS,WORD_TO_STRING(C_PORT,'%u'));

    IF C_MODE<BYTE#4 THEN
      IP4_TO_STRING(IP4:=C_IP);
      CS := CONCAT(CS,' /IP=');
      CS := CONCAT(CS,IP4_TO_STRING.IP4_TO_STRING);
    END_IF;

    ERROR_TIME := MAX(UDINT#200,TIME_TO_UDINT2(TIME_OUT));
    IP_C.TIME_RESET := TRUE;
  END_IF;

  C_ENABLE := IP_C.C_ENABLE AND NOT C_RECONNECT AND NOT NEW_CONNECTION AND IP_C.ERROR = DWORD#0;

  FB_IP_CONNECT.EN_C    := C_ENABLE;
  FB_IP_CONNECT.PARTNER := CS;
  FB_IP_CONNECT();
  C_READY  := FB_IP_CONNECT.VALID;
  C_ERROR  := FB_IP_CONNECT.ERROR;
  C_STATUS := FB_IP_CONNECT.STATUS;
  C_ID     := FB_IP_CONNECT.ID;

  IF C_ENABLE THEN
    IF NOT C_ENABLE_OLD THEN
      DELAY_VALUE := UDINT#50;
    END_IF;
  ELSE
    IF C_ENABLE_OLD THEN
      C_RECONNECT := FALSE;
      DELAY_VALUE := UDINT#50;
    END_IF;
  END_IF;

  C_ENABLE_OLD := C_ENABLE;

  IF C_READY THEN
    IF NOT C_READY_OLD THEN
      IP_C.C_STATE := BYTE#254;
      DELAY_VALUE := UDINT#50;
      IP_C.TIME_RESET := TRUE;

    ELSE
      IP_C.C_STATE := BYTE#255;
    END_IF;
  ELSE
    IF C_READY_OLD THEN
      IP_C.C_STATE := BYTE#1;
    IP_C.MAILBOX[1] := BYTE#0;
    IP_C.MAILBOX[2] := BYTE#0;
    IP_C.MAILBOX[3] := BYTE#0;
      DELAY_VALUE := UDINT#50;

      IF NOT NEW_CONNECTION THEN
        S_ACTIVE := FALSE;
        S_REQ := FALSE;
        S_BUF.SIZE := UINT#0;
      END_IF;
    ELSE
      IP_C.C_STATE := BYTE#000;
    END_IF;
  END_IF;

  C_READY_OLD := C_READY;

  C := 1;
  IF S_BUF.SIZE > UINT#0 THEN
    IF C_READY AND C_ENABLE THEN
      IF S_ACTIVE = FALSE AND IP_C.MAILBOX[2] = BYTE#0 THEN
        S_TOTAL := LIMIT_INT(0,UINT_TO_INT(S_BUF.SIZE),R_E_MAX_SIZE);
        S_CUR_POS  := 0;
        S_CUR_SIZE := 0;
        S_START := TRUE;
        S_ACTIVE := TRUE;
      END_IF;

      IF S_DONE OR S_START THEN

        S_START := FALSE;
        S_CUR_POS := S_CUR_POS + S_CUR_SIZE;
        IF S_TOTAL > S_CUR_POS THEN
          S_CUR_SIZE := S_TOTAL - S_CUR_POS;
          S_CUR_SIZE:=LIMIT_INT(0,S_CUR_SIZE,S_MAX_SIZE);

          C2 := S_CUR_POS;
      C3 := S_CUR_SIZE - 1;
      FOR C := 0 TO C3 DO
            S_BUF_I.BUFFER[C] := S_BUF.BUFFER[C2];
        C2 := C2 + 1;
          END_FOR;
          S_BUF_I.SIZE := INT_TO_UINT(S_CUR_SIZE);
        S_TIME := tx;
          R_TIME := tx;
          S_REQ := TRUE;
          C := 0;
        ELSE
          S_REQ := FALSE;
          S_BUF.SIZE := UINT#0;
          S_ACTIVE := FALSE;
        END_IF;
      END_IF;
    END_IF;
  END_IF;

  FOR C2 := C TO 1 DO
    FB_IP_USEND.REQ    := S_REQ AND C2=1;
    FB_IP_USEND.ID     := C_ID;
    FB_IP_USEND.R_ID   := '';
    FB_IP_USEND.SD_1   := S_BUF_I;
    FB_IP_USEND();
    S_DONE   := FB_IP_USEND.DONE;
    S_ERROR  := FB_IP_USEND.ERROR;
    S_STATUS := FB_IP_USEND.STATUS;
    S_BUF_I  := FB_IP_USEND.SD_1;
  END_FOR;

  FB_IP_URCV.EN_R := C_READY AND NOT S_ACTIVE AND IP_C.MAILBOX[3] = BYTE#0;
  FB_IP_URCV.ID   := C_ID;
  FB_IP_URCV.R_ID := '';
  FB_IP_URCV.RD_1 := R_BUF_I;
  FB_IP_URCV();
  R_NDR    := FB_IP_URCV.NDR;
  R_ERROR  := FB_IP_URCV.ERROR;
  R_STATUS := FB_IP_URCV.STATUS;
  R_BUF_I  := FB_IP_URCV.RD_1;

  IF R_NDR THEN
    IF R_BUF.SIZE >= INT_TO_UINT(R_E_MAX_SIZE) THEN
      R_BUF.SIZE := UINT#0;
      r_status := 254;
    END_IF;

    R_TIME := tx;
    R_COUNT := UINT_TO_INT(R_BUF_I.SIZE);
    R_OFFSET := UINT_TO_INT(R_BUF.SIZE);

    IF (C_MODE AND BYTE#2#0000_0001) = BYTE#1 THEN
      r_offset := 0;
    ELSE
      R_OFFSET := UINT_TO_INT(R_BUF.SIZE);
    END_IF;

    IF R_OFFSET + R_COUNT > R_E_MAX_SIZE THEN
      R_COUNT := R_E_MAX_SIZE - R_OFFSET;
    END_IF;

    C2 := R_OFFSET;
    C3 := R_COUNT - 1;
    FOR C := 0 TO C3 DO
      R_BUF.BUFFER[C2] := R_BUF_I.BUFFER[C];
      C2 := C2 + 1;
    END_FOR;

    R_BUF.SIZE := INT_TO_UINT(R_OFFSET + R_COUNT);
    IP_C.MAILBOX[1] := USINT_TO_BYTE(BYTE_TO_USINT(IP_C.MAILBOX[1]) + USINT#1);
    IF IP_C.MAILBOX[1] = BYTE#0 THEN IP_C.MAILBOX[1] := BYTE#1; END_IF;

  END_IF;

  IF IP_C.TIME_RESET THEN
    IP_C.TIME_RESET := FALSE;
    C_RECONNECT_COUNT := 0;
    C_TIME := tx;
    S_TIME := tx;
    R_TIME := tx;

    ERROR_CON := BYTE#0;
    ERROR_SND := BYTE#0;
    ERROR_RCV := BYTE#0;
  END_IF;

  IF IP_C.R_OBSERVE = FALSE OR s_active THEN
      R_TIME := tx;
  END_IF;

  C_RECONNECT := FALSE;

  IF ERROR_CON = BYTE#0 THEN
    IF C_ERROR THEN
    IF C_STATUS = 16#31 THEN
      ERROR_CON := BYTE#253;
    ELSE
      ERROR_CON := INT_TO_BYTE(C_STATUS);
    END_IF;
    ELSIF TX - C_TIME > ERROR_TIME AND C_ENABLE AND NOT C_READY AND C_MODE < BYTE#2 THEN
      IF C_RECONNECT_COUNT >= 3 THEN
        ERROR_CON := BYTE#255;
      ELSE
        C_TIME := TX;
        C_RECONNECT_COUNT := C_RECONNECT_COUNT + 1;
        C_RECONNECT := TRUE;

      END_IF;
    END_IF;
  END_IF;

  IF ERROR_SND = BYTE#0 THEN
    IF S_ERROR AND S_STATUS <> 16#65 THEN
      ERROR_SND := INT_TO_BYTE(S_STATUS);
    ELSIF TX - S_TIME > ERROR_TIME AND S_ACTIVE THEN
      ERROR_SND := BYTE#255;
    END_IF;
  END_IF;

  IF ERROR_RCV = BYTE#0 THEN
    IF R_ERROR AND (R_STATUS <> 16#33) AND (R_STATUS <> 16#31) AND (R_STATUS <> 16#65) THEN
      ERROR_RCV := INT_TO_BYTE(R_STATUS);
    ELSIF TX - R_TIME > ERROR_TIME AND C_READY AND IP_C.R_OBSERVE THEN
      ERROR_RCV := BYTE#255;
    END_IF;
  END_IF;

  IP_C.ERROR := DWORD_OF_BYTE(ERROR_CON,ERROR_SND,ERROR_RCV,BYTE#0);

END_FUNCTION_BLOCK

PROGRAM program0
	VAR
		IP :	DWORD;
    PORT :	WORD;
    TIME_OUT :	TIME;
    IP_C :	oscat_IP_C;
    S_BUF :	oscat_NETWORK_BUFFER;
    R_BUF :	oscat_NETWORK_BUFFER;

		func_block : IP_CONTROL_Block;
	END_VAR
	func_block.IP := IP;
	func_block.PORT := PORT;
	func_block.TIME_OUT := TIME_OUT;
	func_block.IP_C := IP_C;
	func_block.S_BUF := S_BUF;
	func_block.R_BUF := R_BUF;

	func_block();
  IP_C  := func_block.IP_C;
	S_BUF  := func_block.S_BUF;
	R_BUF  := func_block.R_BUF;

END_PROGRAM

CONFIGURATION Config0
	RESOURCE Res0 ON PLC
		TASK task0(INTERVAL := T#20ms,PRIORITY := 0);
		PROGRAM instance0 WITH task0 : program0;
	END_RESOURCE
END_CONFIGURATION

(* ---- IP_CONTROL2.ST ---- *)
FUNCTION_BLOCK IP_CONTROL2

  VAR

  END_VAR

  VAR_EXTERNAL

  END_VAR

  VAR

  END_VAR

  VAR
    T_PLC_MS :	T_PLC_MS;
    IP4_TO_STRING :	IP4_TO_STRING;
    FB_IP_CONNECT :	IP_CONNECT;
    FB_IP_URCV :	IP_URCV;
    FB_IP_USEND :	IP_USEND;
  END_VAR

  VAR_INPUT
    IP :	DWORD;
    PORT :	WORD;
    TIME_OUT :	TIME;
  END_VAR

  VAR_IN_OUT
    IP_C :	oscat_IP_C;
    S_BUF :	oscat_NETWORK_BUFFER_SHORT;
    R_BUF :	oscat_NETWORK_BUFFER_SHORT;
  END_VAR

  VAR
    C_TIME :	UDINT;
    S_TIME :	UDINT;
    R_TIME :	UDINT;
    C_ENABLE :	BOOL;
    C_IP :	DWORD;
    C_PORT :	WORD;
    C_MODE :	BYTE;
    C_ERROR :	BOOL;
    C_STATUS :	INT;
    C_ID :	INT;
    C_RECONNECT :	BOOL;
    C_RECONNECT_COUNT :	INT;
    S_DONE :	BOOL;
    S_ERROR :	BOOL;
    S_STATUS :	INT;
    S_ACTIVE :	BOOL;
    R_NDR :	BOOL;
    R_ERROR :	BOOL;
    R_STATUS :	INT;
    NEW_CONNECTION :	BOOL;
    C_ENABLE_OLD :	BOOL;
    C_READY :	BOOL;
    C_READY_OLD :	BOOL;
    DELAY_STOP :	UDINT;
    DELAY :	UDINT;
    DELAY_VALUE :	UDINT;
    C :	INT;
    C2 :	INT;
    CS :	oscat_STRING50;
    TX :	UDINT;
    ERROR_TIME :	UDINT;
    ERROR_CON :	BYTE;
    ERROR_SND :	BYTE;
    ERROR_RCV :	BYTE;
  END_VAR

  T_PLC_MS();
  TX := T_PLC_MS.T_PLC_MS;

  IF (TX - DELAY < DELAY_VALUE) THEN
    IF IP_C.C_STATE <> BYTE#1 AND IP_C.C_STATE <> BYTE#254 THEN
    RETURN;
    END_IF;
  END_IF;
  DELAY := TX;

  IF C_ENABLE AND DELAY_VALUE > UDINT#00 THEN
    IF (TX - DELAY_STOP > UDINT#1000) THEN
      DELAY_VALUE := UDINT#00;

    END_IF;
  ELSE
    DELAY_STOP := TX;
  END_IF;

  IF IP_C.C_PORT = WORD#00 THEN
    IP_C.C_PORT := PORT;
  END_IF;
  IF IP_C.C_IP=DWORD#00 AND IP_C.C_MODE<BYTE#4 THEN
    IP_C.C_IP := IP;
  END_IF;

  NEW_CONNECTION := C_IP <> IP_C.C_IP OR C_MODE <> IP_C.C_MODE OR C_PORT <> IP_C.C_PORT;

  IF IP_C.C_ENABLE AND NOT C_READY AND NEW_CONNECTION THEN

    C_IP   := IP_C.C_IP;
    C_MODE := IP_C.C_MODE;
    C_PORT := IP_C.C_PORT;

    CS := SEL_STRING((C_MODE AND BYTE#1) = BYTE#1,'','/UDP ');
    CS := CONCAT(CS,SEL_STRING(C_MODE<BYTE#2,'/PASSIVE','/ACTIVE'));
    CS := CONCAT(CS,' /PORT=');
    CS := CONCAT(CS,WORD_TO_STRING(C_PORT,'%u'));

    IF C_MODE<BYTE#4 THEN
      IP4_TO_STRING(IP4:=C_IP);
      CS := CONCAT(CS,' /IP=');
      CS := CONCAT(CS,IP4_TO_STRING.IP4_TO_STRING);
    END_IF;

    ERROR_TIME := MAX(UDINT#200,TIME_TO_UDINT2(TIME_OUT));
    IP_C.TIME_RESET := TRUE;
  END_IF;

  C_ENABLE := IP_C.C_ENABLE AND NOT C_RECONNECT AND NOT NEW_CONNECTION AND IP_C.ERROR = DWORD#0;

  FB_IP_CONNECT.EN_C    := C_ENABLE;
  FB_IP_CONNECT.PARTNER := CS;
  FB_IP_CONNECT();
  C_READY  := FB_IP_CONNECT.VALID;
  C_ERROR  := FB_IP_CONNECT.ERROR;
  C_STATUS := FB_IP_CONNECT.STATUS;
  C_ID     := FB_IP_CONNECT.ID;

  IF C_ENABLE THEN
    IF NOT C_ENABLE_OLD THEN
      DELAY_VALUE := UDINT#50;
    END_IF;
  ELSE
    IF C_ENABLE_OLD THEN
      C_RECONNECT := FALSE;
      DELAY_VALUE := UDINT#50;
    END_IF;
  END_IF;

  C_ENABLE_OLD := C_ENABLE;

  IF C_READY THEN
    IF NOT C_READY_OLD THEN
      IP_C.C_STATE := BYTE#254;
      DELAY_VALUE := UDINT#50;
      IP_C.TIME_RESET := TRUE;
    ELSE
      IP_C.C_STATE := BYTE#255;
    END_IF;
  ELSE
    IF C_READY_OLD THEN
      IP_C.C_STATE := BYTE#1;
    IP_C.MAILBOX[1] := BYTE#0;
    IP_C.MAILBOX[2] := BYTE#0;
    IP_C.MAILBOX[3] := BYTE#0;
      DELAY_VALUE := UDINT#50;

      IF NOT NEW_CONNECTION THEN
        S_ACTIVE := FALSE;
        S_BUF.SIZE := UINT#0;
      END_IF;
    ELSE
      IP_C.C_STATE := BYTE#000;
    END_IF;
  END_IF;

  C_READY_OLD := C_READY;
  C := 1;
  IF S_BUF.SIZE > UINT#0 THEN
    IF C_READY AND C_ENABLE AND S_ACTIVE = FALSE AND IP_C.MAILBOX[2] = BYTE#0 THEN
      S_ACTIVE := TRUE;
      S_TIME := tx;
      R_TIME := tx;
      C := 0;
    END_IF;
  END_IF;

  FOR C2 := C TO 1 DO
    FB_IP_USEND.REQ    := S_ACTIVE AND C2=1;
    FB_IP_USEND.ID     := C_ID;
    FB_IP_USEND.R_ID   := '';
    FB_IP_USEND.SD_1   := S_BUF;
    FB_IP_USEND();
    S_DONE   := FB_IP_USEND.DONE;
    S_ERROR  := FB_IP_USEND.ERROR;
    S_STATUS := FB_IP_USEND.STATUS;
    S_BUF    := FB_IP_USEND.SD_1;
  END_FOR;

  IF S_DONE THEN
      S_ACTIVE := FALSE;
      S_BUF.SIZE := UINT#0;
  END_IF;

  FB_IP_URCV.EN_R := C_READY AND NOT S_ACTIVE AND IP_C.MAILBOX[3] = BYTE#0;
  FB_IP_URCV.ID   := C_ID;
  FB_IP_URCV.R_ID := '';
  FB_IP_URCV.RD_1 := R_BUF;
  FB_IP_URCV();
  R_NDR    := FB_IP_URCV.NDR;
  R_ERROR  := FB_IP_URCV.ERROR;
  R_STATUS := FB_IP_URCV.STATUS;
  R_BUF    := FB_IP_URCV.RD_1;

  IF R_NDR THEN
      R_TIME := TX;
      IP_C.MAILBOX[1] := USINT_TO_BYTE(BYTE_TO_USINT(IP_C.MAILBOX[1]) + USINT#1);
      IF IP_C.MAILBOX[1] = BYTE#0 THEN IP_C.MAILBOX[1] := BYTE#1; END_IF;
  END_IF;

  IF IP_C.TIME_RESET THEN
    IP_C.TIME_RESET := FALSE;
    C_RECONNECT_COUNT := 0;
    C_TIME := tx;
    S_TIME := tx;
    R_TIME := tx;

    ERROR_CON := BYTE#0;
    ERROR_SND := BYTE#0;
    ERROR_RCV := BYTE#0;
  END_IF;

  IF IP_C.R_OBSERVE = FALSE OR s_active THEN
      R_TIME := tx;
  END_IF;

  C_RECONNECT := FALSE;

  IF ERROR_CON = BYTE#0 THEN
    IF C_ERROR THEN
    IF C_STATUS = 16#31 THEN
      ERROR_CON := BYTE#253;
    ELSE
      ERROR_CON := INT_TO_BYTE(C_STATUS);
    END_IF;
    ELSIF TX - C_TIME > ERROR_TIME AND C_ENABLE AND NOT C_READY AND C_MODE < BYTE#2 THEN
      IF C_RECONNECT_COUNT >= 3 THEN
        ERROR_CON := BYTE#255;
      ELSE
        C_TIME := TX;
        C_RECONNECT_COUNT := C_RECONNECT_COUNT + 1;
        C_RECONNECT := TRUE;
      END_IF;
    END_IF;
  END_IF;

  IF ERROR_SND = BYTE#0 THEN
    IF S_ERROR AND S_STATUS <> 16#65 THEN
      ERROR_SND := INT_TO_BYTE(S_STATUS);
    ELSIF TX - S_TIME > ERROR_TIME AND S_ACTIVE THEN
      ERROR_SND := BYTE#255;
    END_IF;
  END_IF;

  IF ERROR_RCV = BYTE#0 THEN
    IF R_ERROR AND (R_STATUS <> 16#33) AND (R_STATUS <> 16#31) AND (R_STATUS <> 16#65) THEN
      ERROR_RCV := INT_TO_BYTE(R_STATUS);
    ELSIF TX - R_TIME > ERROR_TIME AND C_READY AND IP_C.R_OBSERVE THEN
      ERROR_RCV := BYTE#255;
    END_IF;
  END_IF;

  IP_C.ERROR := DWORD_OF_BYTE(ERROR_CON,ERROR_SND,ERROR_RCV,BYTE#0);

END_FUNCTION_BLOCK

(* ---- IP_FIFO.ST ---- *)
TYPE
  oscat_IP_FIFO128_DATA  : ARRAY [1..128] OF BYTE;
  oscat_Mailbox  : ARRAY [1..16] OF BYTE;

  oscat_IP_FIFO_DATA :
  STRUCT
	X       : oscat_IP_FIFO128_DATA; (* IP_ID FIFO Speicher          *)
	Y       : oscat_IP_FIFO128_DATA; (* IP_ID Z�hler                 *)
	ID      : BYTE;                  (* h�chste vergabene id         *)
	MAX_ID  : BYTE;                  (* maximal Anmeldungen pro ID   *)
    INIT    : BOOL;                  (* Initialisierung durchgef�hrt *)
	EMPTY   : BOOL;                  (* FIFO leer                    *)
	FULL    : BOOL;                  (* FIFO voll                    *)
	TOP     : INT;                   (* maximale anzahl in FIFO      *)
	NW      : INT;                   (* Schreibzeiger                *)
	NR      : INT;                   (* Lesezeiger                   *)
  END_STRUCT;
END_TYPE

TYPE

  oscat_NW_BUF_LONG  : ARRAY [0..4095] OF BYTE;

  oscat_NETWORK_BUFFER :
  STRUCT
    SIZE   : UINT;
    BUFFER : oscat_NW_BUF_LONG;
  END_STRUCT;

END_TYPE

FUNCTION _BYTE_TO_INT:INT
	VAR_INPUT
		IN :	BYTE;
	END_VAR

	_BYTE_TO_INT := USINT_TO_INT(BYTE_TO_USINT(IN));
END_FUNCTION

FUNCTION_BLOCK IP_FIFO_Block

  VAR_IN_OUT
    FIFO :	oscat_IP_FIFO_DATA;
    ID :	BYTE;
    STATE :	BYTE;
  END_VAR

  VAR
    tmp :	INT;
  END_VAR

  IF NOT FIFO.INIT THEN
    FIFO.INIT		:= TRUE;
    FIFO.NW		:= 1;
    FIFO.NR		:= 1;
    FIFO.EMPTY	:= TRUE;
    FIFO.FULL		:= FALSE;
    FIFO.TOP		:= 128;
    FIFO.MAX_ID	:= BYTE#1;
  END_IF;

  IF ID = BYTE#00 THEN
    IF FIFO.ID < INT_TO_BYTE(FIFO.TOP) THEN
      ID := USINT_TO_BYTE(BYTE_TO_USINT(FIFO.ID) + USINT#1);
      FIFO.ID := ID ;

    ELSIF STATE < BYTE#200 THEN
      STATE := BYTE#255;
    RETURN;
    END_IF;
  END_IF;

  IF STATE = BYTE#1 AND NOT FIFO.FULL THEN
    tmp := _BYTE_TO_INT(ID);
    IF FIFO.Y[tmp] < FIFO.MAX_ID THEN
      FIFO.Y[tmp] := USINT_TO_BYTE(BYTE_TO_USINT(FIFO.Y[tmp]) + USINT#1);
      tmp := FIFO.NW;
      FIFO.X[tmp] := ID;
      IF FIFO.NW = FIFO.TOP THEN FIFO.NW := 1; ELSE FIFO.NW := FIFO.NW + 1; END_IF;
      FIFO.FULL := FIFO.NW = FIFO.NR;
    FIFO.EMPTY := FALSE;
      STATE := BYTE#2;
    END_IF;
  END_IF;

  IF STATE = BYTE#2 AND NOT FIFO.EMPTY THEN
    tmp := FIFO.NR;
    IF ID = FIFO.X[tmp] THEN
      STATE := BYTE#3;
    END_IF;
  END_IF;

  IF STATE = BYTE#4 AND NOT FIFO.EMPTY THEN

    tmp := FIFO.NR;
    IF ID = FIFO.X[tmp] THEN
      tmp := _BYTE_TO_INT(ID);
      FIFO.Y[tmp] := USINT_TO_BYTE(BYTE_TO_USINT(FIFO.Y[tmp]) - USINT#1);

      IF FIFO.NR = FIFO.TOP THEN FIFO.NR := 1; ELSE FIFO.NR := FIFO.NR + 1; END_IF;
      FIFO.EMPTY := FIFO.NR = FIFO.NW;
    FIFO.FULL := FALSE;
    END_IF;
    STATE := BYTE#5;
  END_IF;

END_FUNCTION_BLOCK

PROGRAM program0
	VAR
		FIFO :	oscat_IP_FIFO_DATA;
    ID :	BYTE;
    STATE :	BYTE;

		func_block : IP_FIFO_Block;
	END_VAR
	func_block.FIFO := FIFO;
	func_block.ID := ID;
  func_block.STATE := STATE;

	func_block();
  FIFO  := func_block.FIFO;
	ID  := func_block.ID;
  STATE  := func_block.STATE;
END_PROGRAM

CONFIGURATION Config0
	RESOURCE Res0 ON PLC
		TASK task0(INTERVAL := T#20ms,PRIORITY := 0);
		PROGRAM instance0 WITH task0 : program0;
	END_RESOURCE
END_CONFIGURATION

(* ---- IRTRANS_DECODE.ST ---- *)
FUNCTION_BLOCK CHR_TO_STRING_Block
	VAR_INPUT
		C :	BYTE;
	END_VAR

	VAR_OUTPUT
		CHR_TO_STRING :	STRING;
	END_VAR

	CHR_TO_STRING := BYTE_TO_STRING(C);

END_FUNCTION_BLOCK

TYPE

  oscat_NW_BUF_SHORT : ARRAY [0..1407] OF BYTE;
  oscat_NW_BUF_LONG  : ARRAY [0..4095] OF BYTE;

  oscat_NETWORK_BUFFER_SHORT :
  STRUCT
    SIZE   : UINT;
    BUFFER : oscat_NW_BUF_SHORT;
  END_STRUCT;

  oscat_NETWORK_BUFFER :
  STRUCT
    SIZE   : UINT;
    BUFFER : oscat_NW_BUF_LONG;
  END_STRUCT;

END_TYPE

TYPE
  oscat_IP_FIFO128_DATA  : ARRAY [1..128] OF BYTE;
  oscat_Mailbox  : ARRAY [1..16] OF BYTE;

  oscat_IP_FIFO_DATA :
  STRUCT
	X       : oscat_IP_FIFO128_DATA; (* IP_ID FIFO Speicher          *)
	Y       : oscat_IP_FIFO128_DATA; (* IP_ID Z�hler                 *)
	ID      : BYTE;                  (* h�chste vergabene id         *)
	MAX_ID  : BYTE;                  (* maximal Anmeldungen pro ID   *)
    INIT    : BOOL;                  (* Initialisierung durchgef�hrt *)
	EMPTY   : BOOL;                  (* FIFO leer                    *)
	FULL    : BOOL;                  (* FIFO voll                    *)
	TOP     : INT;                   (* maximale anzahl in FIFO      *)
	NW      : INT;                   (* Schreibzeiger                *)
	NR      : INT;                   (* Lesezeiger                   *)
  END_STRUCT;

  oscat_IP_C:
  STRUCT
  	C_MODE:			BYTE;          		(*W Mode: TCP/UCP AKTIV/PASSIV                               *)
	C_PORT:         WORD;          		(*W Portnummer                                               *)
	C_IP:           DWORD;         		(*W IP-Adresse gepackt wwxxyyzz = www.xxx.yyy.zzz            *)
    C_STATE:        BYTE;          		(*R Verbindungsstatus ON/OFF + Flanke ON/OFF                 *)
	C_ENABLE:       BOOL;          		(*W Freigabe f�r Connect                                     *)
    R_OBSERVE:      BOOL;          		(*W Empfang ueberwachen                                      *)
    TIME_RESET:     BOOL;          		(*W Alle Timer ruecksetzen                                   *)
	ERROR:          DWORD;         		(*R vvwwxxyy (vv = CON_ERROR, ww = SEN_ERROR, xx = REC_ERROR *)
    FIFO:           oscat_IP_FIFO_DATA; (*I IP FIFO Struktur                                         *)
	MAILBOX:		oscat_Mailbox;		(*I Mailbox: Datenbereich f�r Bausteindatenaustausch         *)
  END_STRUCT;
END_TYPE

FUNCTION_BLOCK IRTRANS_DECODE_Block

	VAR_OUTPUT
		CMD :	BOOL;
		DEV :	STRING;
		KEY :	STRING;
		ERROR :	BOOL;
	END_VAR

	VAR_IN_OUT
		IP_C :	oscat_IP_C;
		R_BUF :	oscat_NETWORK_BUFFER;
	END_VAR

	VAR
		i :	INT;
		stop :	INT;
		received_string :	STRING;
		char :	STRING;
		CHR_TO_STRING :	CHR_TO_STRING_Block;
		z :	BYTE;
	END_VAR

	i := UINT_TO_INT(R_BUF.SIZE);
	IF i >= 5 AND (i <= 82) AND IP_C.MAILBOX[1] <> z THEN
		error := TRUE;
		i := i - 1;

		IF R_BUF.BUFFER[i] <> BYTE#10 THEN RETURN; END_IF;
		i := i - 1;
		IF R_BUF.BUFFER[i] <> BYTE#13 THEN RETURN; END_IF;
		i := i - 1;

		stop := 0;
		received_string := '';

		WHILE stop <= i DO
			CHR_TO_STRING(C:=R_BUF.BUFFER[stop]);
			char := CHR_TO_STRING.CHR_TO_STRING;
			received_string := CONCAT(received_string,char);
			stop := stop + INT#1;
		END_WHILE;

		stop := FIND(received_string,',');
		IF stop > 0 AND stop - 1 < i THEN
			DEV := LEFT(received_string,stop - 1);
			key := RIGHT(received_string,i - stop + 1);
			IF LEN(DEV) = 0 OR LEN(key) = 0 THEN RETURN; END_IF;
			cmd := TRUE;
			error := FALSE;
		END_IF;
	ELSE
		cmd := FALSE;
		error := FALSE;
	END_IF;

	z := IP_C.MAILBOX[1];

END_FUNCTION_BLOCK

PROGRAM program0
	VAR
		IP_C :	oscat_IP_C;
		R_BUF :	oscat_NETWORK_BUFFER;
		CMD :	BOOL;
		DEV :	STRING;
		KEY :	STRING;
		ERROR :	BOOL;

		func_block : IRTRANS_DECODE_Block;
	END_VAR
	func_block.IP_C := IP_C;
	func_block.R_BUF := R_BUF;

	func_block();
	IP_C  := func_block.IP_C;
	R_BUF  := func_block.R_BUF;
	CMD  := func_block.CMD;
	DEV  := func_block.DEV;
	KEY  := func_block.KEY;
	ERROR  := func_block.ERROR;

END_PROGRAM

CONFIGURATION Config0

  	RESOURCE Res0 ON PLC
    	TASK task0(INTERVAL := T#20ms,PRIORITY := 0);
    	PROGRAM instance0 WITH task0 : program0;
  	END_RESOURCE

END_CONFIGURATION

(* ---- IRTRANS_RCV_1.ST ---- *)
FUNCTION_BLOCK IRTRANS_RCV_1_Block

	VAR_INPUT
		CMD :	BOOL;
		DEV_CODE :	STRING;
		KEY_CODE :	STRING;
	END_VAR

	VAR_OUTPUT
		Q :	BOOL;
	END_VAR

	VAR_IN_OUT
		DEV :	STRING;
		KEY :	STRING;
	END_VAR

	Q := cmd AND EQ_STRING(dev_code,dev) AND EQ_STRING(key_code,key);

END_FUNCTION_BLOCK

PROGRAM program0
	VAR
		CMD :	BOOL;
		DEV :	STRING;
		KEY :	STRING;
		DEV_CODE :	STRING;
		KEY_CODE :	STRING;
		Q :	BOOL;

		func_block : IRTRANS_RCV_1_Block;
	END_VAR
	func_block.CMD := CMD;
	func_block.DEV := DEV;
	func_block.KEY := KEY;
	func_block.DEV_CODE := DEV_CODE;
	func_block.KEY_CODE := KEY_CODE;

	func_block();
	DEV  := func_block.DEV;
	KEY  := func_block.KEY;
	Q  := func_block.Q;

END_PROGRAM

CONFIGURATION Config0

  	RESOURCE Res0 ON PLC
    	TASK task0(INTERVAL := T#20ms,PRIORITY := 0);
    	PROGRAM instance0 WITH task0 : program0;
  	END_RESOURCE

END_CONFIGURATION

(* ---- IRTRANS_RCV_4.ST ---- *)
FUNCTION_BLOCK IRTRANS_RCV_4_Block

	VAR_INPUT
		CMD :	BOOL;
	END_VAR

	VAR_IN_OUT
		DEV :	STRING;
		KEY :	STRING;
	END_VAR

	VAR_INPUT
		DEV_CODE :	STRING;
		KEY_CODE_0 :	STRING;
		KEY_CODE_1 :	STRING;
		KEY_CODE_2 :	STRING;
		KEY_CODE_3 :	STRING;
	END_VAR

	VAR_OUTPUT
		Q0 :	BOOL;
		Q1 :	BOOL;
		Q2 :	BOOL;
		Q3 :	BOOL;
	END_VAR

	VAR
		decode :	BOOL;
	END_VAR

	decode := cmd AND EQ_STRING(dev_code,dev);

	Q0 := EQ_STRING(key,key_code_0) AND decode;
	Q1 := EQ_STRING(key,key_code_1) AND decode;
	Q2 := EQ_STRING(key,key_code_2) AND decode;
	Q3 := EQ_STRING(key,key_code_3) AND decode;

END_FUNCTION_BLOCK

PROGRAM program0
	VAR
		CMD :	BOOL;
		DEV :	STRING;
		KEY :	STRING;
		DEV_CODE :	STRING;
		KEY_CODE_0 :	STRING;
		KEY_CODE_1 :	STRING;
		KEY_CODE_2 :	STRING;
		KEY_CODE_3 :	STRING;
		Q0 :	BOOL;
		Q1 :	BOOL;
		Q2 :	BOOL;
		Q3 :	BOOL;

		func_block : IRTRANS_RCV_4_Block;
	END_VAR
	func_block.CMD := CMD;
	func_block.DEV := DEV;
	func_block.KEY := KEY;
	func_block.DEV_CODE := DEV_CODE;
	func_block.KEY_CODE_0 := KEY_CODE_0;
	func_block.KEY_CODE_1 := KEY_CODE_1;
	func_block.KEY_CODE_2 := KEY_CODE_2;
	func_block.KEY_CODE_3 := KEY_CODE_3;

	func_block();
	DEV  := func_block.DEV;
	KEY  := func_block.KEY;
	Q0  := func_block.Q0;
	Q1  := func_block.Q1;
	Q2  := func_block.Q2;
	Q3  := func_block.Q3;

END_PROGRAM

CONFIGURATION Config0

  	RESOURCE Res0 ON PLC
    	TASK task0(INTERVAL := T#20ms,PRIORITY := 0);
    	PROGRAM instance0 WITH task0 : program0;
  	END_RESOURCE

END_CONFIGURATION

(* ---- IRTRANS_RCV_8.ST ---- *)
FUNCTION_BLOCK IRTRANS_RCV_8_Block

	VAR_INPUT
		CMD :	BOOL;
	END_VAR

	VAR_IN_OUT
		DEV :	STRING;
		KEY :	STRING;
	END_VAR

	VAR_INPUT
		DEV_CODE :	STRING;
		KEY_CODE_0 :	STRING;
		KEY_CODE_1 :	STRING;
		KEY_CODE_2 :	STRING;
		KEY_CODE_3 :	STRING;
		KEY_CODE_4 :	STRING;
		KEY_CODE_5 :	STRING;
		KEY_CODE_6 :	STRING;
		KEY_CODE_7 :	STRING;
	END_VAR

	VAR_OUTPUT
		Q0 :	BOOL;
		Q1 :	BOOL;
		Q2 :	BOOL;
		Q3 :	BOOL;
		Q4 :	BOOL;
		Q5 :	BOOL;
		Q6 :	BOOL;
		Q7 :	BOOL;
	END_VAR

	VAR
		decode :	BOOL;
	END_VAR

	decode := cmd AND EQ_STRING(dev_code,dev);

	Q0 := EQ_STRING(key,key_code_0) AND decode;
	Q1 := EQ_STRING(key,key_code_1) AND decode;
	Q2 := EQ_STRING(key,key_code_2) AND decode;
	Q3 := EQ_STRING(key,key_code_3) AND decode;
	Q4 := EQ_STRING(key,key_code_4) AND decode;
	Q5 := EQ_STRING(key,key_code_5) AND decode;
	Q6 := EQ_STRING(key,key_code_6) AND decode;
	Q7 := EQ_STRING(key,key_code_7) AND decode;

END_FUNCTION_BLOCK

PROGRAM program0
	VAR
		CMD :	BOOL;
		DEV :	STRING;
		KEY :	STRING;
		DEV_CODE :	STRING;
		KEY_CODE_0 :	STRING;
		KEY_CODE_1 :	STRING;
		KEY_CODE_2 :	STRING;
		KEY_CODE_3 :	STRING;
		KEY_CODE_4 :	STRING;
		KEY_CODE_5 :	STRING;
		KEY_CODE_6 :	STRING;
		KEY_CODE_7 :	STRING;
		Q0 :	BOOL;
		Q1 :	BOOL;
		Q2 :	BOOL;
		Q3 :	BOOL;
		Q4 :	BOOL;
		Q5 :	BOOL;
		Q6 :	BOOL;
		Q7 :	BOOL;

		func_block : IRTRANS_RCV_8_Block;
	END_VAR
	func_block.CMD := CMD;
	func_block.DEV := DEV;
	func_block.KEY := KEY;
	func_block.DEV_CODE := DEV_CODE;
	func_block.KEY_CODE_0 := KEY_CODE_0;
	func_block.KEY_CODE_1 := KEY_CODE_1;
	func_block.KEY_CODE_2 := KEY_CODE_2;
	func_block.KEY_CODE_3 := KEY_CODE_3;
	func_block.KEY_CODE_4 := KEY_CODE_4;
	func_block.KEY_CODE_5 := KEY_CODE_5;
	func_block.KEY_CODE_6 := KEY_CODE_6;
	func_block.KEY_CODE_7 := KEY_CODE_7;

	func_block();
	DEV  := func_block.DEV;
	KEY  := func_block.KEY;
	Q0  := func_block.Q0;
	Q1  := func_block.Q1;
	Q2  := func_block.Q2;
	Q3  := func_block.Q3;
	Q4  := func_block.Q4;
	Q5  := func_block.Q5;
	Q6  := func_block.Q6;
	Q7  := func_block.Q7;

END_PROGRAM

CONFIGURATION Config0

  	RESOURCE Res0 ON PLC
    	TASK task0(INTERVAL := T#20ms,PRIORITY := 0);
    	PROGRAM instance0 WITH task0 : program0;
  	END_RESOURCE

END_CONFIGURATION

(* ---- IRTRANS_SERVER.ST ---- *)
TYPE

  oscat_NW_BUF_SHORT : ARRAY [0..1407] OF BYTE;
  oscat_NW_BUF_LONG  : ARRAY [0..4095] OF BYTE;

  oscat_NETWORK_BUFFER_SHORT :
  STRUCT
    SIZE   : UINT;
    BUFFER : oscat_NW_BUF_SHORT;
  END_STRUCT;

  oscat_NETWORK_BUFFER :
  STRUCT
    SIZE   : UINT;
    BUFFER : oscat_NW_BUF_LONG;
  END_STRUCT;

END_TYPE

TYPE
  oscat_IP_FIFO128_DATA  : ARRAY [1..128] OF BYTE;
  oscat_Mailbox  : ARRAY [1..16] OF BYTE;

  oscat_IP_FIFO_DATA :
  STRUCT
	X       : oscat_IP_FIFO128_DATA; (* IP_ID FIFO Speicher          *)
	Y       : oscat_IP_FIFO128_DATA; (* IP_ID Z�hler                 *)
	ID      : BYTE;                  (* h�chste vergabene id         *)
	MAX_ID  : BYTE;                  (* maximal Anmeldungen pro ID   *)
    INIT    : BOOL;                  (* Initialisierung durchgef�hrt *)
	EMPTY   : BOOL;                  (* FIFO leer                    *)
	FULL    : BOOL;                  (* FIFO voll                    *)
	TOP     : INT;                   (* maximale anzahl in FIFO      *)
	NW      : INT;                   (* Schreibzeiger                *)
	NR      : INT;                   (* Lesezeiger                   *)
  END_STRUCT;

  oscat_IP_C:
  STRUCT
  	C_MODE:			BYTE;          		(*W Mode: TCP/UCP AKTIV/PASSIV                               *)
	C_PORT:         WORD;          		(*W Portnummer                                               *)
	C_IP:           DWORD;         		(*W IP-Adresse gepackt wwxxyyzz = www.xxx.yyy.zzz            *)
    C_STATE:        BYTE;          		(*R Verbindungsstatus ON/OFF + Flanke ON/OFF                 *)
	C_ENABLE:       BOOL;          		(*W Freigabe f�r Connect                                     *)
    R_OBSERVE:      BOOL;          		(*W Empfang ueberwachen                                      *)
    TIME_RESET:     BOOL;          		(*W Alle Timer ruecksetzen                                   *)
	ERROR:          DWORD;         		(*R vvwwxxyy (vv = CON_ERROR, ww = SEN_ERROR, xx = REC_ERROR *)
    FIFO:           oscat_IP_FIFO_DATA; (*I IP FIFO Struktur                                         *)
	MAILBOX:		oscat_Mailbox;		(*I Mailbox: Datenbereich f�r Bausteindatenaustausch         *)
  END_STRUCT;
END_TYPE

FUNCTION_BLOCK IRTRANS_SERVER_Block

	VAR_INPUT
		UDP_TCP :	BOOL;
	END_VAR

	VAR_OUTPUT
		S_ENABLE :	BOOL;
		R_ENABLE :	BOOL;
		ERROR :	DWORD;
	END_VAR

	VAR_IN_OUT
		IP_C :	oscat_IP_C;
		S_BUF :	oscat_NETWORK_BUFFER;
		R_BUF :	oscat_NETWORK_BUFFER;
	END_VAR

	VAR
		t :	TON;
	END_VAR

	IF NOT IP_C.C_ENABLE THEN
		IP_C.C_PORT := WORD#0;
		IP_C.C_IP := DWORD#00;
		IP_C.C_MODE := SEL(UDP_TCP,BYTE#5,BYTE#4);
		IP_C.C_ENABLE := TRUE;
		IP_C.R_OBSERVE := FALSE;
		IP_C.TIME_RESET := TRUE;
		S_BUF.SIZE := UINT#0;
		R_BUF.SIZE := UINT#0;
	END_IF;

	R_ENABLE := IP_C.C_STATE > BYTE#127;
	S_ENABLE := R_ENABLE AND (IP_C.MAILBOX[1] > BYTE#0 OR IP_C.C_MODE <> BYTE#5);
	ERROR := IP_C.ERROR;

	t(IN:= IP_C.ERROR > DWORD#0, PT:=T#5s);
	IF t.Q THEN
		IP_C.TIME_RESET := TRUE;
	END_IF;

END_FUNCTION_BLOCK

PROGRAM program0
	VAR
		UDP_TCP :	BOOL;
		S_ENABLE :	BOOL;
		R_ENABLE :	BOOL;
		ERROR :	DWORD;
		IP_C :	oscat_IP_C;
		S_BUF :	oscat_NETWORK_BUFFER;
		R_BUF :	oscat_NETWORK_BUFFER;

		func_block : IRTRANS_SERVER_Block;
	END_VAR
	func_block.UDP_TCP := UDP_TCP;
	func_block.IP_C := IP_C;
	func_block.S_BUF := S_BUF;
	func_block.R_BUF := R_BUF;

	func_block();
	S_ENABLE  := func_block.S_ENABLE;
	R_ENABLE  := func_block.R_ENABLE;
	ERROR  := func_block.ERROR;
	IP_C  := func_block.IP_C;
	S_BUF  := func_block.S_BUF;
	R_BUF  := func_block.R_BUF;

END_PROGRAM

CONFIGURATION Config0

  	RESOURCE Res0 ON PLC
    	TASK task0(INTERVAL := T#20ms,PRIORITY := 0);
    	PROGRAM instance0 WITH task0 : program0;
  	END_RESOURCE

END_CONFIGURATION

(* ---- IS_CC.ST ---- *)
FUNCTION_BLOCK IS_CC_Block

	VAR_INPUT
		STR :	STRING;
		CMP :	STRING;
	END_VAR

	VAR_OUTPUT
		IS_CC :	BOOL;
	END_VAR

	VAR
		L :	INT;
		pos :	INT;
		temp :	STRING;
	END_VAR

	L := LEN(str);
	FOR pos := 1 TO L DO
		temp := MID(str,1,pos);
		IF FIND(CMP,temp) = 0 THEN
			IS_CC := FALSE;
			RETURN;
		END_IF;
	END_FOR;
	IS_CC := L > 0;

END_FUNCTION_BLOCK

PROGRAM program0

	VAR
		STR :	STRING;
		CMP :	STRING;

		IS_CC :	BOOL;

		func_block : IS_CC_Block;
	END_VAR
	func_block.STR := STR;
	func_block.CMP := CMP;
	func_block();
	IS_CC := func_block.IS_CC;

END_PROGRAM

CONFIGURATION Config0

	RESOURCE Res0 ON PLC
		TASK task0(INTERVAL := T#20ms,PRIORITY := 0);
		PROGRAM instance0 WITH task0 : program0;
	END_RESOURCE

END_CONFIGURATION

(* ---- IS_IP4.ST ---- *)
FUNCTION_BLOCK IS_IP4

	VAR_INPUT
		STR :	STRING;
	END_VAR

	VAR_OUTPUT
		IS_IP4 :	BOOL;
	END_VAR

	VAR
		COUNT_CHAR :	COUNT_CHAR;
	END_VAR

	COUNT_CHAR(STR:=str,CHR:=BYTE#46);
	IS_IP4 := COUNT_CHAR.COUNT_CHAR = 3;

END_FUNCTION_BLOCK

(* ---- IS_LOWER.ST ---- *)
FUNCTION_BLOCK IS_LOWER

VAR_INPUT
	STR :	STRING;
END_VAR

VAR_OUTPUT
	IS_LOWER :	BOOL;
END_VAR

VAR
	pos :	INT;
	I :	INT;
END_VAR

I := LEN(str);
FOR pos := 1 TO I DO
	IF NOT ISC_LOWER(INT_TO_BYTE(GET_CHAR(str,pos))) THEN
		IS_LOWER := FALSE;
		RETURN;
	END_IF;
END_FOR;
IS_LOWER := I>0;

END_FUNCTION_BLOCK
